(* IEC 61131-3 sources: IRIS-Project/LASAL CONTROL SOFTWARE/LasalProject_2025_09_25/Runtime/%LASALAPPDATA%/Runtime/Library/Loader/Source/code (part 3) *)

  IF SramdiskNotWrittenAtPowerDown() THEN
		DEBUGLOG0("%010d error: sramdisk was not written at power-down");
    _s_ram_hptr^.DataValid$UINT := 0;
    sramErrorCode := EC_SRAMDISK_NOT_WRITTEN_AT_POWER_DOWN;
    LogSramError();
  END_IF;

	IF isRamfileDatUsed THEN
		// Das RAMFILE.DAT auf pRamFile einlesen
		IF SramLoadFile() <> 0 THEN
			_s_ram_hptr^.DataValid$UINT := 0;
			sramErrorCode := EC_LOADFILE_ERR;
			LogSramError();
		ELSIF IsVortex() = FALSE & WasRemoveableMediaChanged() THEN
			DEBUGLOG0("%010d error: detected media change, ramfile.dat not usable, marking sram as invalid");
			_s_ram_hptr^.DataValid$UINT := 0;
		END_IF;
	END_IF;

  fDoNotReportErrors := 0;
  IF GetSramReorgFlag() & ((_s_ram_hptr^.DataValid AND 16#FF000000) = 16#80000000) THEN
    // Wenn das Reorg-Flag im DataValid Feld gesetzt ist, dann heißt das, daß
    // ein Reorg Vorgang unterbrochen wurde, nachdem eine File Kopie angelegt
    // wurde. In so einem Fall wird keine Fehlermeldung generiert.
    fDoNotReportErrors := 1;
  END_IF;

	IF GetSramReorgFlag() THEN
		fReorgSram := 1;
	END_IF;
	wasValid := CHK_S_RAM(fDoNotReportErrors);
	IF GetSramReorgFlag() THEN
		IF wasValid THEN

			// gültigen SRAM Inhalt auf Files kopieren
			rc := MakeSramKopie(#errCode);
			IF rc = 0 THEN

				// Der SRAM Inhalt befindet jetzt als Kopie in den Files.
				// Es wird jetzt als ungültig gekennzeichnet und durch den Aufruf von CHK_S_RAM
				// wird das SRAM noch einmal mit 0 initialisiert.
				DEBUGLOG0("%010d MakeSramKopie succeeded, marking sram as invalid");

				_s_ram_hptr^.DataValid$UINT := 0;
        // Das Reorg-Flag setzen. Wenn dieses Flag gesetz ist, dann heisst das, daß
        // das SRAM zwar ungültig ist, aber eine gültige Kopie im File existiert.
        // In diesem Fall (ungültige SRAM, gültige Kopie im File) wird kein SRAM
        // Fehler gemeldet.
        _s_ram_hptr^.DataValid := (_s_ram_hptr^.DataValid AND 16#00FFFFFF) OR 16#80000000;

        // Der folgende Aufruf von CHK_S_RAM bewirkt, daß das SRAM neu initilisiert
        // wird (weil DataValud 0 ist).
				fReorgSram := 1;
				CHK_S_RAM(fDoNotReportErrors := 1);
        // Reorg-Flag muss hier noch einmal gesetzt werden, da CHK_S_RAM den
        // ganzen Header auf 0 setzt.
        _s_ram_hptr^.DataValid := (_s_ram_hptr^.DataValid AND 16#00FFFFFF) OR 16#80000000;

			ELSE
				DEBUGLOG2("%010d MakeSramKopie failed, rc=%d, errCode = 0x%X" , rc$UDINT, errCode$UDINT);
			END_IF;

		//ELSIF !!WasRemoveableMediaChanged() THEN
    ELSE
			_s_ram_hptr^.DataValid$UINT := 0;
            // Der folgende Aufruf von CHK_S_RAM bewirkt, daß das SRAM neu initilisiert
            // wird (weil DataValid 0 ist). Das ist notwendig, damit in der MAT die
			// durch SRAM_MARKMemory belegten Bereiche wieder freigegeben werden.
			// (SRAM_MARKMemory wurde in CHK_S_RAM aufgerufen, um die vorhandenen
			// SRAM Einträge als belegt zu markieren).
			fReorgSram := 1;
			CHK_S_RAM(fDoNotReportErrors := 1);

			// Das SRAM war ungültig, durch das Setzen des Flags fReorgSram wird
			// versucht, auf Daten von einer früheren Kopie zurückzugreifen.
			fReorgSram := 1;
			DEBUGLOG0("%010d MakeSramKopie: no copy created, because sram is not valid");
		END_IF;
	END_IF;

	CLEAR_LASTENTRY();

END_FUNCTION

//------------------------------------------------------------------------
// S-Ram Initialisieren und ggf alte formate konvertieren (aus active.dat)
//-------------------------------------------------------------------------
// Bei aufruf hat das BS schon in  "_S_RAM_Hptr"  einen pointer auf den S-Ram-Descriptor
// Descriptor eingetragen (oder auch nicht. ein altes system hat dort 0 stehen
//
// Logik : a) _S_RAM_Hptr hat einen gültigen pointer.
//				Wenn der eintrag genutzte länge > 0 ist gelten diese daten
//				Wenn der eintrag genutzte länge = 0 ist, suchen wir eine Active.dat
//
// 06.03.04
// wenn C-IPC konvertieren auf neues format
// es stehen nur noch die Daten im Ram der Rest ist in einem File
// so sparen wir pro eintrag 12 Byte !!!
//
//

FUNCTION S_RAM_INIT

VAR_OUTPUT
	ret_code 		: CONFSTATES;
END_VAR

VAR
	ActiveDatHandle  :DINT;
	DateiKopf     : DatKopf;
	OneRecord     : Eintrag;
	RecNr		  : UDINT;
	I			  : DINT;
	PtChar		  : ^CHAR;
	PtxNextRAM	  : ^XRamCell;
	ptxRamHead	  : ^XRAMHDR;
	RelAdress	  :  UDINT;
  formatChanged : BOOL;
  initCnt : UDINT;
	gotMemory : BOOL;
END_VAR

  if !!hasSram then
    ret_code:=C_OK;
    return;
  end_if;

  CONVERT_SRAM();

	// das erstellen wir automatisch
  if _rtosversion > 16#537 then
    if LSLFILE_IsInstalled then
      // Das Direktory für die File Daten erstellen
      OS_FILE_CREATEDIR("C:\FData");
    end_if;
  end_if;

  ret_code:=C_OK;
  initCnt := 0;
Brutal_start:
  initCnt += 1;

//---------------------------------------
// Wenn Neues BS ist der Ptr ungleich 0
//---------------------------------------

  IF _S_RAM_Hptr <> 0 then      // Diesen Pointer gibt es seit a.m mit pranz und gradl am 2.2.2002 vergangenheitsbewältigung gemacht hat

    if (_S_RAM_Hptr^.DataLength <= maxSramSize) then
      SRAM_STARTUP(_S_RAM_Hptr^.DataLength , 1);
    else
      SRAM_STARTUP(maxSramSize, 1);  // SRAM begrenzen
    end_if;

    //------------------------------------------------------
    // wenn jungfräulich, test ob alte active.dat vorhanden
    //------------------------------------------------------
    IF _S_RAM_Hptr^.UsedData = 0 then

      //-- Neues _SRAM Löschen ---

      // Der Aufruf dieser Funktion bewirkt, dass auch bei gelöschtem Sram
      // das File sernum.dat, wo die Seriennummer gespeichert ist, erstellt wird.
      WasRemoveableMediaChanged();

      RelAdress:=InitXramBlockEx(#gotMemory);
      IF gotMemory THEN
        ptxRamHead:= _S_RAM_Hptr^.DataStart+RelAdress;
        PtxNextRam:=#ptxRamHead^.aData[0];

        // active.dat nur möglich wenn filesystem vorhanden

        IF (LSLFILE_IsInstalled) THEN

          ActiveDatHandle:=OS_FILE_OPEN("c:\active.dat",0,16#000);

          // das file ist gefunden -> konvertieren
          IF ActiveDatHandle > 0 THEN
            OS_FILE_READ(ActiveDatHandle, #DateiKopf.signi[0], sizeof(DateiKopf));
            IF DateiKopf.NrRec <> 0 then  // #FA wenn keine eintraege ende  (gibt es auch)
              FOR RecNr:= 0 to DateiKopf.NrRec -1 do
                // -- GUID LESEN
                OS_FILE_READ(ActiveDatHandle,#OneRecord.myguid[0],sizeof(Eintrag.myguid));
                // -- NAMEN LESEN

                PtCHar:=#OneRecord.Name[0];
                FOR I:= 0 to SIZEOF(Eintrag.Name) -1 do
                  OS_FILE_READ(ActiveDatHandle,PtCHar,1);
                  if PtChar^ =0 then
                    GOTO GOTNAME;
                  elsif PtChar^ = '.' then
                    PtChar^:=0;
                  end_if;
                  PtCHar+=1;
                END_FOR;

                // ERROR NAME TO LONG !!!!

                ret_code:=C_OUTOF_NEAR;
                OS_FILE_CLOSE(ActiveDatHandle);
                GOTO	Brutal_ende;

              //...........................
              // Der Name ist eingelesen !
              //...........................

              GOTNAME:

                // wenn block voll, neuen block erzeugen & Verkettung herstellen

                if ptxRamHead^.udEntries = X_RAM_CELLS	then
                  RelAdress:=IniNewRamBlock(PtxNextRam);
                  If Reladress <> 0 then
                    ptxRamHead:= _S_RAM_Hptr^.DataStart+RelAdress;
                    PtxNextRam:=#ptxRamHead^.aData[0];
                    // Kein platz mehr im RAM !!!
                  else
                    ret_code:=C_OUTOF_NEAR;
                    OS_FILE_CLOSE(ActiveDatHandle);
                    GOTO	Brutal_ende;
                  end_if;
                end_if;

                // Daten und Sizeof daten lesen

                OneRecord.CRC:=CRC32(#OneRecord.Name[0]);

                OS_FILE_READ(ActiveDatHandle,#OneRecord.Data,2*4);

                // Wenn Len > 0 dann ist es eine RAMEX falls es eine RAMEX mit 0 ist
                // kommt das später beim Instanzieren dran

                IF OneRecord.Len <> 0 then
                  RelAdress$UDINT:= (SRAM_GetMemory(OneRecord.Len$UDINT))$UDINT;
                  If Reladress <> 0 then

                    PtxNextRam^.udType:=IsXram$UDINT+RelAdress$UDINT;
                    OS_FILE_READ(ActiveDatHandle,_S_RAM_Hptr^.DataStart+RelAdress,OneRecord.Len$UDINT);
                    // in the data HIGH Part is the real length
                    // in the lo part the allocated length
                    OneRecord.Data$UDINT := OneRecord.Len$UDINT SHL 16;
                    OneRecord.Data$UDINT := OneRecord.Data$UDINT OR  SRAM_GET_ALLOCATED(OneRecord.Len$UDINT);
                  end_if;

                ELSE
                  PtxNextRam^.udType:= 0;
                END_IF;

                PtxNextRam^.udCRC32:=OneRecord.CRC;
                PtxNextRam^.udData$UDINT:=OneRecord.Data$UDINT;
                PtxNextRam^.udChk$UDINT:=OneRecord.Data$UDINT+OneRecord.CRC+(PtxNextRam^.udType$UDINT AND 16#00ffFFFF);
                PtxNextRam^.udType:=PtxNextRam^.udType or RamValid;  // VALID RAM LOCATION

                ptxNextRam+=SIZEOF(xRamCell);
                ptxRamHead^.udEntries+=1;
                ptxRamHead^.udChk:=NOT ptxRamHead^.udEntries;

              END_FOR;
            END_IF;
            OS_FILE_CLOSE(ActiveDatHandle);
            S_RAM_INIT_I();

          // keine active.dat vorhanden  und neues system und dateisystemvorhanden .
          //--> Speicher Initialisieren
          ELSE
            S_RAM_INIT_I();
          END_IF;

        // Kein filesystem vorhanden & keine daten: jungfräulich, initialisieren
        // oder das alte Format konvertieren !
        // muss eigentlich Eine 386 sein ??

        ELSE
          // #FA
          // wir versuchen die alten daten auch zu konvertieren aber nur einmal
          if aRamHdr.udEntries <> 0 then
            if aRamHdr.udEntries = NOT aRamHdr.udChk then
              if aRamHdr.udEntries < 1000 then // sicherheit
                // schleife für die konvertierung bilden !!!
                for RecNr:=0 to (aRamHdr.udEntries-1) do

                  // wenn block voll, neuen block erzeugen & Verkettung herstellen
                  if ptxRamHead^.udEntries = X_RAM_CELLS	then
                    RelAdress:=IniNewRamBlock(PtxNextRam);
                    If Reladress <> 0 then
                      ptxRamHead:= _S_RAM_Hptr^.DataStart+RelAdress;
                      PtxNextRam:=#ptxRamHead^.aData[0];
                    // Kein platz mehr im RAM !!!
                    else
                      ret_code:=C_OUTOF_NEAR;
                      GOTO	Brutal_ende;
                    end_if;
                  end_if;

                  // check if chk is o.k.
                  if aRamHdr.aData[RecNr].udChk = aRamHdr.aData[RecNr].udCRC32 + aRamHdr.aData[RecNr].udData then
                    PtxNextRam^.udCRC32:=aRamHdr.aData[RecNr].udCRC32;
                    PtxNextRam^.udData$UDINT:=aRamHdr.aData[RecNr].udData;
                    PtxNextRam^.udChk$UDINT:=aRamHdr.aData[RecNr].udChk;

                    PtxNextRam^.udType:=PtxNextRam^.udType or RamValid;  // VALID RAM LOCATION

                    ptxNextRam+=SIZEOF(xRamCell);
                    ptxRamHead^.udEntries+=1;
                    ptxRamHead^.udChk:=NOT ptxRamHead^.udEntries;
                  end_if;

                end_for;
              end_if;
            end_if;
            aRamHdr.udEntries :=0;
            aRamHdr.udChk :=0;
          end_if;

          S_RAM_INIT_I();
        END_IF;
      ELSE // gotMemory
        IF !!isRamfileDatUsed THEN
          // Bei SRAM Format 1 muss auf jeden Fall der xRamHdr Platz haben
          LDR_outOfSramMem := TRUE;
        END_IF;

        S_RAM_INIT_I();
      END_IF;

    //--- ES SIND DATEN VORHANDEN, TESTEN !!! ---

    ELSE
      S_RAM_INIT_I();
    END_IF;

  //------------------------------------
  // ALTES FORMAT (kein Ptr auf ram vorhanden)
  //------------------------------------
  else
    ret_code:=C_OUTOF_NEAR;
  END_IF;
Brutal_ende:

  IF loaderRamexError THEN
    IF isSramNewOrCleared THEN
      DEBUGLOG0("%010d-resetting sram content due to a detected new or cleared sram");
    ELSE
      DEBUGLOG0("%010d-resetting sram content due to a detected error");
    END_IF;
    LDR_outOfSramMem := FALSE;
    _s_ram_hptr^.UsedData := 0;
    _s_ram_hptr^.DataStart^.udEntries := 0;
    _s_ram_hptr^.DataStart^.udChk:=NOT _s_ram_hptr^.DataStart^.udEntries;
    IF GetRamfileDatUsedFlag(#formatChanged) THEN
      _s_ram_hptr^.DataValid := 0x20001;
    ELSE
      _s_ram_hptr^.DataValid := 0x00001;
    END_IF;
    IF pRamFile THEN
      pRamFile^.udEntries :=  0;
      pRamFile^.uiChange  :=  16#1234;	// änderung eintragen wir speicher hier gleich
    END_IF;
    SramSaveFile();

    // DS2589, 02.02.182, 9.5.2016:
    // Eine möglicherweise von früher noch vorhandene Sram-Kopie (vom Reorganisieren)
    // wird gelöscht, damit im Fall einer gesetzten SRAM_CONTINUE_ON_ERROR Umgebungsvariable
    // das Sram mit den Init-Werten und nicht mit den Werten aus der Kopie initialisiert wird.
    DeleteSramKopie();

    IF (!!bSramContinueOnError & !!isSramNewOrCleared) | (initCnt > 1) THEN
      ret_code:=C_OUTOF_NEAR;
    ELSIF formatChanged THEN
      // Wenn das Format geändert wurde, dann muss noch einmal initialisiert
      // werden (es ist z.B. die Größe der MAT vom Format abhängig).
      loaderRamexError := 0;
      GOTO Brutal_start;
    END_IF;
  END_IF;

END_FUNCTION

// Löscht im alten Format in der letzten Zelle des ersten Blocks den im Element
// udType (in den untersten 20 Bits) gespeicherten Merker für die letzte gefundene
// Ramzelle. Dieser Merker wird von der Funktion Find_sRam_I zum Zwischenspeichern
// des Block-Index und Zell-Offsets der zuletzt gefundenen Zelle verwendet.
// Damit wird die Suche schneller, wenn Find_sRam_I nicht jedesmal von vorne
// zu suchen beginnt, sondern dort wo sie den letzten Eintrag gefunden hat.
//
// Im neuen Format (mit ramfile.dat) wird dieser Merker nicht verwendet.
FUNCTION CLEAR_LASTENTRY
VAR
  pRamCell : ^XRamCell;
END_VAR;

  IF (_S_RAM_Hptr^.DataValid SHR 16) < 2 &  _s_ram_hptr^.DataLength >= SIZEOF(XRAMHDR) THEN
    // altes Format
    pRamCell := #_S_RAM_Hptr^.DataStart^.aData[X_RAM_CELLS];
    pRamCell^.udType := pRamCell^.udType AND 16#FFF0_0000;
  END_IF;

END_FUNCTION

// loescht alle Einträge
FUNCTION ClearEntrys

	pRamFile^.udEntries   := 0;
	pRamFile^.CRC32       := 0;
	pRamFile^.pLastEntry  := 0;

END_FUNCTION

#define READ_COMPLETE_RAMFILEDAT

// Wenn das Sram im RAM liegt mit einem Backup auf SD Karte (Edge-CPUs),
// dann wird in dieser Funktion der Sram-Inhalt auf die SD Karte gesichert.
FUNCTION FlushSramToDisk
VAR
  pSrd : ^OS_SRAMDISK;
END_VAR

  OS_CILGet("SRAMDISK", #pSrd$void);
  IF (pSrd <> NIL) & (pSrd^.udVersion >= 2) THEN
    SRAMDISK_COMMIT(pSrd);
#ifdef _LSL_TARGETARCH_X86
    // SA26191,DS2087: Workaround für einen OS-Fehler bei ETVEdge Plattformen:
    // Interrupts sind nach Aufruf von SRAMDISK_COMMIT gesperrt, wenn fullCopyAtPowerdown gesetzt ist.
    // Die Interrupts werden hier wieder freigegeben.
    IF _RtOSVersion < 16#9000 THEN
      STI();
    END_IF;
#endif
  END_IF;

END_FUNCTION

// funktion schreibt daten auf Flash falls verson C-IPC +
// die Version > 2 ist und sich auch was geändert hat !! in diesem File
FUNCTION GLOBAL SramSaveFile
VAR
	Handle : DINT;
	CRC32  : UDINT;
	aXFileHdr_Hdr : XFILEHDR_HDR;
	pCopy  : ^XFILEHDR;
	rc     : UDINT;
	bytes2Write	 : UDINT;
	bytes2Read   : UDINT;
  allocSize : UDINT;
  att : UDINT;
END_VAR

  if !!hasSram then
    return;
  end_if;

	// test auf C-IPC
	if isRamfileDatUsed then
 	  // test auf pointer vorhanden und version groesser 1
	  if (_S_RAM_Hptr <> NIL) & ((_S_RAM_Hptr^.DataValid shr 16) > 1) then

      if pRamFile^.uichange <> 16#1234 then
        // Wenn keine Änderung war und noch kein RamFile.dat existiert (neuer CIPC),
        // dann wird pRamFile^.uichange auf 16#1234 gesetzt. Dadurch wird das Anlegen
        // eines (leeren) RamFile.dat erzwungen.
        Handle:=OS_FILE_OPEN("c:\RamFile.dat",0,16#000);	// read-only
        if handle >= 0 then
          OS_FILE_CLOSE(handle);
        else
          pRamFile^.uichange := 16#1234;
        end_if;
      end_if;

      // test ob auch sich was geändert hat
      if pRamFile^.uichange = 16#1234 then
        // Ab 1.1.27 wird das SRAM bei jedem Start reorganisiert.
        // Die pRamFile Struktur wird immer neu aufgebaut, d.h. uichange hat
        // dann immer den Wert 16#1234 weil immer Änderungen gemacht werden.
        // Jetzt kann es aber sein, daß die Struktur gleich geblieben ist (wenn sich
        // die Checksumme und udEntries nicht geändert hat). Wenn das der Fall ist, dann
        // wird uichange auf 0 gesetzt, damit das RAMFILE.DAT nicht unnötigerweise
        // neu erstellt wird.

        // Checksumme rechnen
  #ifdef READ_COMPLETE_RAMFILEDAT
        CRC32 := CALC_RAMFILE_DAT_CRC(pRamFile);
  #else
        CRC32:=CRC32_Buffer(#pRamFile^.aData,pRamFile^.udEntries * SIZEOF(XFileCell));
  #endif
        // Checksumme aus dem File einlesen und vergleichen
        handle := OS_FILE_OPEN("c:\RamFile.dat", 0, 0);		// 0 = read only
        IF handle > 0 THEN
          rc := OS_FILE_READ(handle, #aXFileHdr_Hdr, SIZEOF(aXFileHdr_Hdr));
          IF rc = SIZEOF(XFileHdr_Hdr) THEN
            IF (aXFileHdr_Hdr.CRC32 = CRC32) & (aXFileHdr_Hdr.udEntries = pRamFile^.udEntries) THEN
              pRamFile^.uichange := 0;
              DEBUGLOG2("%010d-SramSaveFile: no need to write to ramfile.dat (crc32=0x%08X and udEntries=%d are still the same)", CRC32, pRamFile^.udEntries);
            END_IF;
          END_IF;
          OS_FILE_CLOSE(handle);
        END_IF;
      end_if;

      if pRamFile^.uichange = 16#1234 then

        pRamFile^.CRC32 := CRC32;

				// RAMFILE.DAT auf RAMFILE.BAK kopieren
        Handle:=OS_FILE_OPEN("c:\RamFile.dat",0,16#000);
	      if handle >= 0 then
          allocSize := XFILEHDR.adata + X_FILE_CELLS_2 * SIZEOF(XFileCell);
     			pCopy := (_alloc_resize_LDR(allocSize))$^XFILEHDR;
		      if pCopy <> NIL then
						bytes2Read := allocSize;
	     			rc := OS_FILE_READ(Handle, pCopy, bytes2Read);
		        OS_FILE_CLOSE(handle);
						if rc < 0 then
							DEBUGLOG2("%010d-SramSaveFile: error reading ramfile.dat, bytes2read=%d, rc=%d", bytes2read, rc);
						else
		          handle:=OS_FILE_OPEN("c:\RamFile.bak",2,ATT_CREATE);
							if handle >= 0 then
								bytes2Write := rc;
			 					rc := FileWrite(handle, pCopy, bytes2Write)$UDINT;
								if rc <> bytes2Write then
									DEBUGLOG2("%010d-SramSaveFile: error writing ramfile.bak, bytes2write=%d, rc=%d", bytes2Write, rc);
								else
									DEBUGLOG1("%010d-SramSaveFile: ramfile.dat copied into ramfile.bak (%d bytes)", rc);
								end_if;
				 				OS_FILE_CLOSE(handle);
							else
								DEBUGLOG1("%010d-SramSaveFile: could not open ramfile.bak, rc=%d", handle$UDINT);
							end_if;
	          end_if;
	     		  _free(pCopy);
					else
					  DEBUGLOG1("%010d-SramSaveFile: could not allocate enough memory (%d)", allocSize$UDINT);
		        OS_FILE_CLOSE(handle);
	        end_if;
	   		end_if;

        // den Inhalt von pRamFile ins File RAMFILE.DAT schreiben
        if pRamFile^.udEntries > X_FILE_CELLS then
          bytes2Write := XFILEHDR.adata + X_FILE_CELLS_2 * SIZEOF(XFileCell);
        else
          bytes2Write := XFILEHDR.adata + X_FILE_CELLS * SIZEOF(XFileCell);
        end_if;
        if bytes2Write <> LDR_allocated_XFileSize then
          att := ATT_CREATE_ALWAYS;
        else
          att := ATT_CREATE;
        end_if;

        handle:=OS_FILE_OPEN("c:\RamFile.dat", 2, att);
        if Handle >= 0 then
          rc := FileWrite(handle, pRamFile, bytes2Write)$UDINT;
          if rc <> bytes2Write then
            DEBUGLOG2("%010d-SramSaveFile: error writing ramfile.dat, bytes2write=%d, rc=%d", bytes2Write, rc);
            SramError();
          else
            DEBUGLOG3("%010d-SramSaveFile: data written to ramfile.dat (%d bytes, crc32=0x%X), udEntries=%d", rc, pRamFile^.CRC32, pRamFile^.udEntries);
            // Wenn das Sram im RAM liegt mit einem Backup auf SD Karte (Edge-CPUs),
            // dann wird nach dem Ändern der ramfile.dat der Sram-Inhalt auf die SD Karte
            // geschrieben. Damit ist ramfile.dat und Sram konsistent, auch für den Fall dass
            // beim Abschalten das Sram nicht mehr auf die SD Karte geschriben wird.
            FlushSramToDisk();
            pRamFile^.uichange := 0;
          end_if;
          OS_FILE_CLOSE(handle);
        else
          DEBUGLOG1("%010d-SramSaveFile: could not open ramfile.dat, rc=%d", handle$UDINT);
          Trace_ERR("SAVE OF RamFile not possible (Disk full??)");
          LSLCLI_LoaderTracePrint("SAVE OF RamFile not possible (Disk full??)", 12);
          SramError();
        end_if;

        // ramfile.bak ungültig machen, nachdem ramfile.dat erstellt worden ist
        InvalidateRamfileBak();

      end_if;
    end_if;
	end_if;
END_FUNCTION

// ------------------------------------------
//   laden des File von C-IPC in Speicher
// ------------------------------------------
// das file ist 192k /4 Byte (je Eintrag im S-RAM) * 12 byte (je Eintrag im File)
// groß = 576 k Byte
// die RamEx bleibt so wie alt
// udCRC32    (4 Byte)
// udType     (4 Byte)
// udpRelSram (4 Byte)

FUNCTION SramLoadFile
VAR_OUTPUT
	result : UDINT;
END_VAR
VAR
	Handle : DINT;
	CRC32  : UDINT;
	rc     : UDINT;
	bytes2Read   : UDINT;
	fileSize   : UDINT;
  udEntries_file  : UDINT;
  nCellsAlloc : UDINT;
  allocSize : UDINT;
END_VAR
  result := 16#FFFFFFFF;

  // Die Anzahl der benötigten Zellen ist erst nach dem Lesen des Ramfile.dat
  // bekannt, da aber nachfolgender Code davon ausgeht, dass pRamfile <> NIL ist, wird
  // hier einmal mit X_FILE_CELLS allokiert. Ggf. wird das dann noch vergrößert.
  nCellsAlloc := X_FILE_CELLS;
  allocSize := XFILEHDR.adata + nCellsAlloc * SIZEOF(XFileCell);
	pRamFile := _alloc_resize_LDR(allocSize)$^XFILEHDR;
  if pRamFile <> NIL then
    LDR_allocated_XFileCells := nCellsAlloc;
    LDR_allocated_XFileSize := allocSize;
    ClearEntrys();
  end_if;

  Handle := OS_FILE_OPEN("c:\RamFile.dat",0,0);
  if Handle < 0 then
    DEBUGLOG1("%010d-SramLoadFile: could not open ramfile.dat, rc=%d", handle$UDINT);
    SramError();
    return;
  end_if;
  rc := OS_FILE_READ(Handle, #udEntries_file, SIZEOF(udEntries_file));
  if rc <> SIZEOF(udEntries_file) then
    DEBUGLOG1("%010d-SramLoadFile: could not read udEntries_file from ramfile.dat, rc=%d", rc);
    SramError();
    return;
  end_if;
  OS_FILE_CLOSE(handle);

  if udEntries_file > X_FILE_CELLS & pRamFile <> NIL then
    nCellsAlloc := X_FILE_CELLS_2;
    allocSize := XFILEHDR.adata + nCellsAlloc * SIZEOF(XFileCell);
   	pRamFile := _realloc_LDR(pRamFile, allocSize)$^XFILEHDR;
  end_if;

  if pRamFile <> NIL then
    LDR_allocated_XFileCells := nCellsAlloc;
    LDR_allocated_XFileSize := allocSize;

    ClearEntrys();

    // try to open file
    Handle:=OS_FILE_OPEN("c:\RamFile.dat",0,0);
	  if Handle > 0 then
	 // file ist da laden
#ifdef READ_COMPLETE_RAMFILEDAT
			bytes2Read := allocSize;
			rc := OS_FILE_READ(Handle, pRamFile, bytes2Read);
#else
			rc := OS_FILE_READ(Handle, pRamFile, SIZEOF(XFILEHDR.udEntries));
      if rc = SIZEOF(XFILEHDR.udEntries) then
			  bytes2Read := XFILEHDR.adata + pRamFile^.udEntries * SIZEOF(XFileCell) - SIZEOF(XFILEHDR.udEntries);
			  rc := OS_FILE_READ(Handle, pRamFile + SIZEOF(XFILEHDR.udEntries), bytes2Read);
      end_if;
#endif
	    OS_FILE_CLOSE(handle);
      fileSize := XFILEHDR.adata + pRamFile^.udEntries * SIZEOF(XFileCell);
			if rc < 0 then
				DEBUGLOG1("%010d-SramLoadFile: error reading ramfile.dat, no header information, rc=%d", rc);
				SramError();
			elsif rc <> bytes2Read then
				DEBUGLOG3("%010d-SramLoadFile: error reading ramfile.dat, fileSize=%d, bytes2Read=%d, rc=%d", fileSize, bytes2Read, rc);
				SramError();
			else
	      // file im Speicher CRC rechnen
	      pRamFile^.uiChange :=0;				// keine Änderung
	      pRamFile^.pLastEntry :=0;				// und von anfang an
#ifdef READ_COMPLETE_RAMFILEDAT
	      CRC32 := CALC_RAMFILE_DAT_CRC(pRamFile);
#else
	      CRC32:=CRC32_Buffer(#pRamFile^.aData,pRamFile^.udEntries * SIZEOF(XFileCell));
#endif

	      if CRC32 = pRamFile^.CRC32 then
	        // file im speicher CRC = o.k. wir belegen den Speicher
	        if ((pRamFile^.udEntries <> 0) & (pRamFile^.udEntries <= X_FILE_CELLS_2)) then
						DEBUGLOG2("%010d-SramLoadFile: data read from ramfile.dat (%d bytes), udEntries=%d", rc, pRamFile^.udEntries);
	          result:=0;
	        else
						if pRamFile^.udEntries > X_FILE_CELLS_2 then
					  	DEBUGLOG1("%010d-SramLoadFile: invalid udEntries (%08X)", pRamFile^.udEntries);
						  SramError();
						else
							result := 0;
						end_if;
						ClearEntrys(); // 0 oder zu viele einträge
  	      end_if;
	      else
					DEBUGLOG2("%010d-SramLoadFile: invalid crc32 (calc:0x%08X, file:0x%08X)", CRC32, pRamFile^.CRC32);
					// die CRC ist falsch

					Handle := OS_FILE_OPEN("c:\RamFile.er1",2,ATT_CREATE);
					FileWrite(handle,pRamFile, allocSize);
					OS_FILE_CLOSE(handle);

          // wir nehmen das BAK falls vorhanden
          Handle:=OS_FILE_OPEN("c:\RamFile.bak",2,ATT_READ_WRITE);
          if Handle > 0 then
            OS_FILE_CLOSE(handle);
            OS_FILE_DELETE("c:\RamFile.dat");
            OS_FILE_RENAME("c:\RamFile.bak", "c:\RamFile.dat");
            _free(pRamFile);			// wird nochmal gemacht !!
            result:=SramLoadFile();	// rekursion !!
          end_if;
	      end_if;
	    end_if;
	  else
			DEBUGLOG1("%010d-SramLoadFile: could not open ramfile.dat, rc=%d", handle$UDINT);
			SramError();
	  end_if;
  end_if;

	IF result <> 0 THEN
   		DEBUGLOG1("%010d-SramLoadFile failed, rc=%d", result);
	END_IF;

END_FUNCTION

//------------------------------------------------------------------------------
// AlarmSramError
//------------------------------------------------------------------------------
FUNCTION AlarmSramError
VAR_INPUT
  param : DINT;
END_VAR
	IF (pSramAlarmSvrCh = NIL) & ( (OPS.SysState = C_RUNRAM) | (OPS.SysState = C_RUNROM) ) THEN
		_LookUpEmbed_C(SRAMALARM_SVR_NAME, #pSramAlarmSvrCh, NIL);
	END_IF;
	IF pSramAlarmSvrCh <> NIL THEN
		ESI := pSramAlarmSvrCh;
		pSramAlarmSvrCh^.pMeth^.pWr$M_WR_DIRECT(param);
	END_IF;
END_FUNCTION
//------------------------------------------------------------------------------
// SramError
//------------------------------------------------------------------------------
FUNCTION SramError
	IF loaderRamexError = 0 THEN
    IF isSramNewOrCleared THEN
		  TRACE("New or cleared SRAM detected, see c:\sysmsg\event19.log. Resetted SRAM.");
      LSLCLI_LoaderTracePrint("New or cleared SRAM detected, see c:\sysmsg\event19.log. Resetted SRAM.", 12);
    ELSIF bSramContinueOnError THEN
		  TRACE_WARN("Error in SRAM, see c:\sysmsg\event19.log. Resetted SRAM.");
      LSLCLI_LoaderTracePrint("Error in SRAM, see c:\sysmsg\event19.log. Resetted SRAM.", 12);
    ELSE
		  TRACE_WARN("Error in SRAM, see c:\sysmsg\event19.log. Resetted SRAM, project must be restarted");
      LSLCLI_LoaderTracePrint("Error in SRAM, see c:\sysmsg\event19.log. Resetted SRAM, project must be restarted", 12);
    END_IF;
	END_IF;
	loaderRamexError := 1;
END_FUNCTION
//------------------------------------------------------------------------------
// LogSramError
//------------------------------------------------------------------------------
FUNCTION LogSramError
	IF sramErrorCode = 4 THEN
		// Der Fehlercode 4 kommt zustande, wenn ein RAMFILE.DAT mit udEntries = 0
		// vorgefunden wird.
		// pr:
		//	Meiner Meinung nach ist das kein Fehler, daher wird hier keine Meldung
		//  ausgegeben.
		//  Es wird aber trotzdem der Code für die Fehlerbehandlung durchlaufen, weil
		//  ich nicht weiss wie der ganze Assemblercode auf udEntries = 0 reagieren würde.
		RETURN;
	END_IF;
	DEBUGLOG1("%010d-SramError, errorCode=%08X", sramErrorCode);
	IF _S_RAM_Hptr THEN
		DEBUGLOG1("%010d             Version    = %08X" , _S_RAM_Hptr^.Version);
		DEBUGLOG1("%010d             DataStart  = %08X" , _S_RAM_Hptr^.DataStart$UDINT);
		DEBUGLOG1("%010d             DataLength = %08X" , _S_RAM_Hptr^.DataLength);
		DEBUGLOG1("%010d             UsedData   = %08X" , _S_RAM_Hptr^.UsedData);
		DEBUGLOG1("%010d             DataValid  = %08X" , _S_RAM_Hptr^.DataValid);
		IF _S_RAM_Hptr^.DataStart THEN
			DEBUGLOG1("%010d             udEntries  = %08X" , _S_RAM_Hptr^.DataStart^.udEntries);
			DEBUGLOG1("%010d             udChk      = %08X" , _S_RAM_Hptr^.DataStart^.udChk);
		END_IF;
	END_IF;
	SramError();
END_FUNCTION
//------------------------------------------------------------------------------
// LogSramRamexError
//------------------------------------------------------------------------------
FUNCTION __CDECL LogSramRamexError
VAR_INPUT
	pXramCell : ^XRamCell;
END_VAR
	DEBUGLOG1("%010d-RamexError, cellAddr = %08X" , pXramCell$UDINT);
	DEBUGLOG1("%010d             udChk    = %08X" , pXramCell^.udChk);
	DEBUGLOG1("%010d             udCRC32  = %08X" , pXramCell^.udCRC32);
	DEBUGLOG1("%010d             udData   = %08X" , pXramCell^.udData);
	DEBUGLOG1("%010d             udType   = %08X" , pXramCell^.udType);
	SramError();
END_FUNCTION
//------------------------------------------------------------------------------
// LogSramChk
//------------------------------------------------------------------------------
FUNCTION LogSramChk
	DEBUGLOG0("%010d-checking Sram");
END_FUNCTION
//------------------------------------------------------------------------------
// SramCheckerInit
//------------------------------------------------------------------------------
FUNCTION SramCheckerInit
	fileCellChkIdx := 0;
END_FUNCTION

#ifdef CYCLIC_SRAM_CHECK
#define CELLMASK_VALID      0x80000000
#define CELLMASK_USED       0x40000000
#define CELLMASK_CELLTYPE   0x3C000000
#define CELLMASK_RAMEXADR   0x00FFFFFF

#define CELLTYPE_RAM        0x00000000
#define CELLTYPE_RAMEX      0x30000000

FUNCTION SramCheckV1
VAR
  pHdr : ^XRAMHDR;
  sramStart : pVoid;
  sramEnd : pVoid;
  pCellEnd : ^XRamCell;
  pCell : ^XRamCell;
  cellChksum : UDINT;
END_VAR

  sramStart := _S_RAM_Hptr^.dataStart;
  sramEnd := sramStart + _S_RAM_Hptr^.dataLength;
  pHdr := _S_RAM_Hptr^.dataStart;

  WHILE ((pHdr >= sramStart) & (pHdr < sramEnd)) DO

    IF pHdr^.udEntries > X_RAM_CELLS + 1 THEN
  		sramErrorCode := EC_INV_BLK_ENTRIES;
      SramError();
      AlarmSramError(pHdr$DINT);
    END_IF;
    IF (pHdr^.udEntries XOR pHdr^.udChk) <> 16#FFFFffff THEN
  		sramErrorCode := EC_INV_BLK_CHKSUM;
      SramError();
      AlarmSramError(pHdr$DINT);
    END_IF;

    pCell := #pHdr^.aData[0];
    pCellEnd := #pHdr^.aData[pHdr^.udEntries];
    WHILE pCell < pCellEnd DO

      IF pCell^.udType AND CELLMASK_VALID THEN
        IF pCell^.udType AND CELLMASK_CELLTYPE AND CELLTYPE_RAMEX THEN
          cellChksum := pCell^.udData + pCell^.udCRC32 + (pCell^.udType AND CELLMASK_RAMEXADR);
        ELSE
          cellChksum := pCell^.udData + pCell^.udCRC32;
        END_IF;
        IF cellChksum <> pCell^.udChk THEN
      		sramErrorCode := EC_INV_CELL_CHKSUM;
          SramError();
          AlarmSramError(pCell$DINT);
        END_IF;
      END_IF;

      pCell += sizeof(XRamCell);
    END_WHILE;

    IF pCell = #pHdr^.aData[X_RAM_CELLS] THEN
      // Block war zur Gänze gefüllt
      // prüfen, ob die 501. Zelle auf einen weiteren Block zeigt
      cellChksum := pCell^.udData + pCell^.udCRC32;
      IF ((pCell^.udCRC32 = 1954) & (pCell^.udType AND CELLMASK_VALID) & (cellChksum = pCell^.udChk)) THEN
        // in der 501.Zelle ist ein Zeiger auf den nächsten XRam-Block
        pHdr := sramStart + pCell^.udData;
        IF ((pHdr < sramStart) | (pHdr >= sramEnd)) THEN
          // Verkettung ungültig
      		sramErrorCode := EC_INV_BLK_CHAIN;
          SramError();
          AlarmSramError(pCell$DINT);
        END_IF;
      ELSE
        pHdr := NIL;
      END_IF;
    ELSE
      // Block war nur teilweise gefüllt, es handelt sich also um den letzten Block
      pHdr := NIL; // bewirkt Schleifenaabruch
    END_IF;

  END_WHILE;

END_FUNCTION

//------------------------------------------------------------------------------
// SramChecker
//------------------------------------------------------------------------------
FUNCTION GLOBAL SramCheckerCyclic
VAR
	pFileCell 	: ^XFileCell;
	pRamCell	: ^XRamCell;
	quit		: BOOL;
	chkSum		: UDINT;
	fileCellCnt	: UDINT;
END_VAR

	// wenn bereits ein Fehler festgestellt wurde, dann nichts mehr prüfen,
	// damit das Logfile nicht voll wird
	IF loaderRamexError <> 0 THEN
		AlarmSramError(1);	// Alarm immer wieder auslösen
		RETURN;
	END_IF;

 	IF _S_RAM_Hptr = NIL THEN
		RETURN;
	END_IF;

 	IF _S_RAM_Hptr^.DataValid < 2 THEN
    SramCheckV1();
		RETURN;
	END_IF;

 	IF !!isRamfileDatUsed THEN
		RETURN;
	END_IF;

	IF pRamFile^.udEntries = 0 THEN
		RETURN;
	END_IF;

(*
	pr, 7.2.05: ab 1.1.3 wird bei udEntries = 0 kein Sramfehler gemeldet
	IF _S_RAM_Hptr^.dataStart^.udEntries = 0 THEN
		sramErrorCode := 10;
		LogSramError();
		AlarmSramError(1);
		RETURN;
	END_IF;
*)

	IF (_S_RAM_Hptr^.dataStart^.udEntries XOR _S_RAM_Hptr^.dataStart^.udChk) <> 16#FFFFffff THEN
		sramErrorCode := EC_INV_BLK0_CHKSUM2;
		LogSramError();
		AlarmSramError(1);
		RETURN;
	END_IF;

	fileCellCnt := 0;
	quit := FALSE;
	WHILE !!quit DO

		pFileCell := #pRamFile^.aData[fileCellChkIdx];
		IF (pFileCell^.udCRC32 <> 0) & ((pFileCell^.udType AND 16#3C00_0000) = isXram) THEN
			// Ramex Zelle gefunden -> Checksumme prüfen, dann Schleife abbrechen
			pRamCell := _S_RAM_Hptr^.dataStart + pFileCell^.udpRelSram;

			chkSum := (pRamCell^.udType AND 16#00ffFFFF) + pRamCell^.udData + pRamCell^.udCRC32;
			IF chkSum <> pRamCell^.udChk THEN
				LogSramRamexError(pRamCell);
				AlarmSramError(pRamCell$DINT);
				//(0$^UDINT)^ := 0;	// Exception auslösen
			END_IF;

			quit := TRUE;
		END_IF;

		fileCellChkIdx += 1;
		IF fileCellChkIdx >= pRamFile^.udEntries THEN
			// das Ende ist erreicht -> index auf 0, dann Schleife abbrechen
			fileCellChkIdx := 0;
			quit := TRUE;
		END_IF;

		fileCellCnt += 1;
		IF fileCellCnt > 15 THEN
			// max. 15 File-Cells pro Durchlauf prüfen (sonst kann ein RUNTIME Error auftreten !)
			quit := TRUE;
		END_IF;

	END_WHILE;

END_FUNCTION
#endif

#ifdef _LSL_TARGETARCH_ARM
(*
  Überprüft den Inhalt der Sram-V2 Datenstruktur ob diese gültig ist
  und markiert den verwendeten Sram-Speicher in der MAT als belegt.

  Wenn der Sram Inhalt inhalt gültig ist, wird 0 zurückgegeben, sonst
  ein entsprechender Fehlercode.
*)
FUNCTION CHK_S_RAMV2
VAR_OUTPUT
  errCode : UDINT;
END_VAR
VAR
  i : UDINT;
  pXRAMHDR : ^XRAMHDR;
  pXRamCell : ^XRamCell;
  pXFileCell : ^XFileCell;
  ramStart :^XRamHdr;
END_VAR

  errCode := 0;

  IF !!(_S_RAM_Hptr^.DataValid AND 1) THEN
    errCode := EC_NOT_VALID;
    RETURN;
  END_IF;

  // In UsedData ist der Header mit eingerechnet
  IF _S_RAM_Hptr^.UsedData > _S_RAM_Hptr^.DataLength + _S_RAM_Hptr^.DataStart$UDINT - _S_RAM_Hptr$UDINT THEN
    errCode := EC_OUT_OF_SRAM;
    RETURN;
  END_IF;

  pXRAMHDR := _S_RAM_Hptr^.DataStart;
  IF pXRAMHDR^.udChk <> NOT pXRAMHDR^.udEntries THEN
    errCode := EC_INV_BLK0_CHKSUM;
    RETURN;
  END_IF;

  ramStart := _S_RAM_Hptr^.DataStart;

  // alle einträge o.k. jetzt machen wir noch eine Belegung im RAM mit dem mapper

  // *****************************************
  // die ersten 8 byte sind besonders //
  // *****************************************
  SRAM_MARKMemory(NIL, 8); //length: XRAMHDR (udEntries + udChk)

  pXFileCell := #pRamFile^.aData[0];
  FOR i := 1 TO pRamFile^.udEntries DO
    IF pXFileCell^.udCRC32 <> 0 THEN
      IF (pXFileCell^.udType AND 16#3C00_0000) <> ISXRAM THEN
        // normale RAMZelle	einfach speicher reservieren

        SRAM_MARKMemory(pXFileCell^.udpRelSram$^USINT, 4);

      ELSE
        // RAMEx Zelle

        pXRamCell := ramStart + pXFileCell^.udpRelSram;

        // 'XRamCell.udCRC32 = XFileCell.udCRC32' darf nicht geprueft werden weil
        // durch exchdataptr woanders liegen kann

        // CRC pruefen
        IF pXRamCell^.udChk = ((pXRamCell^.udType AND 16#00ffFFFF) +
                               pXRamCell^.udData +
                               pXRamCell^.udCRC32) THEN
          // super o.k. --> reservieren 16 byte block + reservieren Datenblock
          SRAM_MARKMemory(pXFileCell^.udpRelSram$^USINT, sizeof(XRamCell));
          SRAM_MARKMemory((pXRamCell^.udType AND 16#00FF_FFFF)$^USINT, pXRamCell^.udData AND 16#ffff);
        ELSE
          // die Ramex weist Fehler auf
          errCode := EC_INV_XRAMCELL_CHKSUM;
          LogSramRamexError(pXRamCell);

          pXFileCell^.udpRelSram := 0; // ungültig machen neuer speicher anlegen
          pXFileCell^.udCRC32 := 0; // loeschen damit nicht mehr gefunden wird

          pRamFile^.uiChange := 16#1234; // merker das Änderung

          pXRamCell^.udType := 0; // daten auch loaschen
          pXRamCell^.udData := 0; // daten auch loaschen
          pXRamCell^.udCRC32 := 0;
          pXRamCell^.udChk := 1;	 // damit chk sicher falsch ist
        END_IF;
      END_IF;
    END_IF;
    pXFileCell += sizeof(XFileCell);
  END_FOR;

END_FUNCTION

#ifdef _LSL_TARGETARCH_ARM_SUPPORTS_SRAMV1
(*
  Initialisiert das Sram im alten Format mit einem leeren Block.
*)
FUNCTION S_RAMV1_INITIALIZE_WITH_ONE_BLOCK
VAR
	sramSize : UDINT;
END_VAR

  _S_RAM_Hptr^.UsedData := 0;
  _S_RAM_Hptr^.DataValid := _S_RAM_Hptr^.DataValid AND 16#8000_0000; // alles außer Reorg-Flag rücksetzen

  IF _S_RAM_Hptr^.DataLength < maxSramSize THEN
    sramSize := _S_RAM_Hptr^.DataLength;
  ELSE
    sramSize := maxSramSize;
  END_IF;
  SRAM_STARTUP(sramSize, 1); // MAT für die Größe des SRAMs anlegen
  InitXramBlock();

END_FUNCTION
#endif // _LSL_TARGETARCH_ARM_SUPPORTS_SRAMV1

#ifdef _LSL_TARGETARCH_ARM_SUPPORTS_SRAMV1
(*
  Überprüft den Inhalt der Sram-V1 Datenstruktur ob diese gültig ist
  und markiert den verwendeten Sram-Speicher in der MAT als belegt.

  Wenn der Sram Inhalt inhalt gültig ist, wird 0 zurückgegeben, sonst
  ein entsprechender Fehlercode.
*)
FUNCTION CHK_S_RAMV1
VAR_OUTPUT
  errCode : UDINT;
END_VAR
VAR
  i : UDINT;
  pXRAMHDR : ^XRAMHDR;
  pXRamCell : ^XRamCell;
  cellValid : BOOL;
  typeFlags : UDINT;
  len : UDINT;
  ofs : UDINT;
END_VAR

  errCode := 0;

  IF !!(_S_RAM_Hptr^.DataValid AND 1) THEN
    errCode := EC_NOT_VALID;
    RETURN;
  END_IF;

  // In UsedData ist der Header mit eingerechnet
   IF _S_RAM_Hptr^.UsedData > _S_RAM_Hptr^.DataLength + _S_RAM_Hptr^.DataStart$UDINT - _S_RAM_Hptr$UDINT THEN
     errCode := EC_OUT_OF_SRAM;
     RETURN;
   END_IF;

  _S_RAM_Hptr^.DataStart^.aData[X_RAM_CELLS].udType :=
    _S_RAM_Hptr^.DataStart^.aData[X_RAM_CELLS].udType AND 16#80FFffff;  // 16*65535 Entries Total(used for quicksearch)

  //- Header prüfen --
  pXRAMHDR := _S_RAM_Hptr^.DataStart;
  WHILE 1 DO

    IF pXRAMHDR^.udEntries > X_RAM_CELLS THEN
      // more than 500 entries in one list !
      errCode := EC_INV_BLK_ENTRIES;
      RETURN;
    END_IF;
    IF pXRAMHDR^.udEntries <> NOT pXRAMHDR^.udChk THEN
      // CHKSUMME nicht OK
      errCode := EC_INV_BLK_CHKSUM;
      RETURN;
    END_IF;

    IF pXRAMHDR^.udEntries = 0 THEN
      S_RAMV1_INITIALIZE_WITH_ONE_BLOCK();	// #FA kommt vor weil active.dat nur header hat und ekien eintrage
      RETURN;
    END_IF;

    //-- Speicherblock belegen  mit länge eines blockes !
    SRAM_MARKMemory(pXRAMHDR$^USINT - _S_RAM_Hptr^.DataStart$UDINT, SIZEOF(XRAMHDR));

    pXRamCell := #pXRAMHDR^.aData[0];
    i := 0;
    WHILE i < pXRAMHDR^.udEntries DO
      cellValid := TRUE;
      IF (pXRamCell^.udType AND RamValid) = 0 THEN // ValidFlg (Bit 31) Must Be High !
        cellValid := FALSE;
      ELSIF pXRamCell^.udChk <> ((pXRamCell^.udType AND 16#00ffFFFF) +
                                 pXRamCell^.udData + pXRamCell^.udCRC32) THEN
        cellValid := FALSE;
      ELSE
        pXRamCell^.udType := pXRamCell^.udType AND NOT RAMUSED; // Clr Used Bit
        // CHK FOR Xtended Ram
        typeFlags := pXRamCell^.udType AND 16#3C00_0000;
        IF typeFlags <> 0 THEN
          IF typeFlags <> IsXram THEN
            cellValid := FALSE;
          END_IF;
        END_IF;
      END_IF;

      IF cellValid THEN
        len := pXRamCell^.udData AND 16#ffff; // mehr als 16#ffff geht nicht
        ofs := pXRamCell^.udType AND 16#00FF_ffff;
        SRAM_MARKMemory(ofs$^USINT, len);
      ELSE
        //--- contens of cell not valid , mark it as free (unused) --
        pXRamCell^.udType := 0;
        pXRamCell^.udData := 0;
        pXRamCell^.udCRC32 := 0;
        pXRamCell^.udChk := 0;
#ifdef SRAM_REPORT_INVALID_CELL1
        // Wenn ein Fehler bei einer Format-1 Zelle gefunden wird, dann wird standardmäßig
        // der Zelleninhalt auf 0 gesetzt und kein Sram Fehler gemeldet.
        // Warum wird kein Fehler gemeldet ?
        // Es hat einmal eine Loaderversion gegeben, bei der eine Sram-Zelle die noch nie
        // beschrieben wurde (also den Init-Wert aufweist), eine ungültige Chksum hatte.
        // Fürs Projekt hatte das keine neg. Auswirkungen, da die Chksum bereichtigt wurde,
        // sobald die Zelle beschrieben wurde (siehe Änderung in 02.02.102, SA17043).
        // Würde man jetzt bei einer falschen Chksum in einer Zelle einen Sram-Fehler melden
        // und das ganze Sram resettieren, dann könnte bei funktionierenden Applikationen
        // das Sram zurückgesetzt werden.
        errCode := EC_INV_V1_CELL;
        RETURN;
#endif
      END_IF;

      pXRamCell += sizeof(XRamCell);
      i += 1;
    END_WHILE;

    // -- CHK FOR NEXT BLOCK --
    IF i < X_RAM_CELLS THEN
      RETURN;
    END_IF;

    IF (pXRamCell^.udCRC32 <> 1954) | !!(pXRamCell^.udType AND RamValid) |
       (((pXRamCell^.udType AND 16#00ff_FFFF) + pXRamCell^.udData + pXRamCell^.udCRC32) <> pXRamCell^.udChk) THEN
      // Mark Cell 500 As EMPTY
      pXRamCell^.udType := 0;
      pXRamCell^.udData := 0;
      pXRamCell^.udCRC32 := 0;
      pXRamCell^.udChk := 0;
      RETURN;
    END_IF;

    pXRamCell := _S_RAM_Hptr^.DataStart + pXRamCell^.udData;

  END_WHILE;

END_FUNCTION
#endif // _LSL_TARGETARCH_ARM_SUPPORTS_SRAMV1
#endif

//-------------------------------------------
// Inhalt der daten im S-RAM -Prüfen und verwendeten Sram-Speicher in der MAT
// als belegt markieren.
//-------------------------------------------

//  udType:
//
// Bit 31.. 1= VALID  (CHksum is OK)
//     30.. 1= USED   (After Startup, it is conected to an Objekt)

//     29..   0   1    			(3000 0000)
//     28..   0   1
//     27..   0   0
//	   26..   0   0
//			  !   +-- 	RAMEX ; UdData field contains LENGTH of data,
//			  +--- RAM
//     25..   Frei
//	   24..   Frei
//
//	   0-23   Relative Startadress  of datablock if RAMEX

// CHK := udCrc+udData+(udType AND 16#00ffffff)

#ifdef _LSL_TARGETARCH_ARM
FUNCTION CHK_S_RAM
VAR_INPUT
  fDoNotReportErrors : UDINT;
END_VAR
VAR_OUTPUT
  wasValid : UDINT;
END_VAR
VAR
	sramSize : UDINT;
  errCode : UDINT;
END_VAR

  LogSramChk();
  wasValid := 1;
  sramErrorCode := 0;

  IF _S_RAM_Hptr^.DataLength < maxSramSize THEN
    sramSize := _S_RAM_Hptr^.DataLength;
  ELSE
    sramSize := maxSramSize;
  END_IF;
  SRAM_STARTUP(sramSize, 1); // MAT für die Größe des SRAMs anlegen

  IF isRamfileDatUsed & ((_S_RAM_Hptr^.DataValid SHR 16) AND 16#7fff) >= 2 THEN // Bit31 von DataValid ist das Reorg-Flag
    // =========================================================================
    // neue Version (mit ramfile.dat)
    // =========================================================================
    errCode := CHK_S_RAMV2();
    IF errCode <> 0 THEN
      sramErrorCode := errCode;
      wasValid := 0;

      IF errCode < 100 THEN
        IF !!fDoNotReportErrors THEN
          LogSramError();
        END_IF;
        // im file alles auf 0
        pRamFile^.udEntries := 0;
        pRamFile^.CRC32 := 0;
        pRamFile^.pLastEntry := 0;
        pRamFile^.uiChange := 16#1234; // merker das Änderung

        // auch im ram alles auf 0
        _S_RAM_Hptr^.UsedData := 0;
        _S_RAM_Hptr^.DataValid := (_S_RAM_Hptr^.DataValid AND 16#8000_0000) OR 16#0002_0000; // alles außer Reorg-Flag rücksetzen
      // und die anzahl der einträge auch loeschen
        _S_RAM_Hptr^.DataStart^.udEntries := 0;
        _S_RAM_Hptr^.DataStart^.udChk := 16#FFFF_ffff;

        IF _S_RAM_Hptr^.DataLength < maxSramSize THEN
          sramSize := _S_RAM_Hptr^.DataLength;
        ELSE
          sramSize := maxSramSize;
        END_IF;
        SRAM_STARTUP(sramSize, 1); // MAT für die Größe des SRAMs anlegen
        SRAM_MARKMemory(NIL, 8); //length: XRAMHDR (udEntries + udChk)
      END_IF;
    END_IF;

    // RAM allociert und als belegt gemeldet jetzt kommen die Konstruktoren der
    // RAM und RAMEX und wollen sich die Pointer holen
  ELSE
#ifdef _LSL_TARGETARCH_ARM_SUPPORTS_SRAMV1
    // =========================================================================
    // alte Version (ohne ramfile.dat)
    // =========================================================================
    errCode := CHK_S_RAMV1();
    IF errCode <> 0 THEN
      sramErrorCode := errCode;
      wasValid := 0;

      IF !!fDoNotReportErrors THEN
        LogSramError();
      END_IF;

      S_RAMV1_INITIALIZE_WITH_ONE_BLOCK();

    END_IF;
#else
    // altes Sram Format wird nicht unterstützt
    sramErrorCode := EC_UNSUPPORTED_FORMAT_V1;
    wasValid := 0;
    IF !!fDoNotReportErrors THEN
      LogSramError();
    END_IF;
#endif

  END_IF;

  GET_USED_S_RAM();

END_FUNCTION
#else
FUNCTION AWL CHK_S_RAM
VAR_INPUT
 fDoNotReportErrors : UDINT;
END_VAR
VAR_OUTPUT
 wasValid : UDINT;
END_VAR
VAR
 MAX_MEM	:UDINT ;
 RamStart   :^XramHdr;
END_VAR

		//*************************
		CALL		LogSramChk
		//*************************

		L.D			wasValid, 1

//	  SRAM_STARTUP(	16#40000 , 1);

		l.eax		_S_RAM_Hptr
		l.eax		(eax+MRAM_DESCR.DataLength)
		cmp.eax		maxSramSize
		jbe			CHK_S_RAMn
		l.eax		maxSramSize
CHK_S_RAMn
		PUSH		EAX			 // result
		PUSH.D		1
		PUSH.D		EAX 		 // Länge von OS
		CALL		SRAM_STARTUP
		ADD.ESP		2*4
		POP			EAX			 // RESULT

		L.D			MAX_MEM,0

   		L.EDI 		_S_RAM_Hptr
// test ob Ramfile.dat verwendet wird
		cmp.b		isRamfileDatUsed, 0
		je			chk_s_ram1

		l.ecx		(EDI+MRAM_DESCR.DataValid)
		shr.ecx		16
		cmp.ecx		2
		jb			chk_s_ram1			 // alte version

// es ist schon eine neue version
		l.ecx		(EDI+MRAM_DESCR.DataValid)
		and.ecx		1
		//*****
		L.D			sramErrorCode,EC_NOT_VALID
		//*****
		jz			chk_s_ram_error		// not valid

    (*DB1875*)
		l.eax		(EDI+MRAM_DESCR.DataLength)
		l.ecx		(EDI+MRAM_DESCR.UsedData)
    add.eax (EDI+MRAM_DESCR.DataStart)  // Header ist in UsedData mit eingerechnet
    sub.eax EDI
    cmp.ecx eax
		//*****
		L.D			sramErrorCode,5
		//*****
		jg			chk_s_ram_error

   		L.EDI		(EDI+MRAM_DESCR.DataStart)
		L.EAX		(EDI+XRAMHDR.udEntries)
		x.EAX		16#ffffffff
		cmp.EAX		(EDI+XRAMHDR.udChk)
		//*****
		L.D			sramErrorCode,EC_INV_BLK0_CHKSUM
		//*****
		jne			chk_s_ram_error

// alle einträge o.k. jetzt machen wir noch eine Belegung im RAM mit dem mapper
		L.EBX		pRamFile
		l.ECX		(EBX+XFILEHDR.udEntries)

		// pr, 21.1.06:
		//	Hier war eine Abfrage ob XFILEHDR.udEntries 0 ist und ein Jump
		//	auf chk_s_ram_error falls es 0 ist. Im Kommentar steht, daß das
		//  ein Fehler ist, der nicht sein kann.
		//	Wieso soll das ein Fehler sein ?
		//	Meiner Meinung nach ist das ganz normal daß XFILEHDR.udEntries 0 ist
		//  wenn ich ein Projekt ohne RAM- und RAMEX- Zellen habe.
		//	Ich war daher so frei und habe diese Abfrage einfach auskommentiert.
		//*****
		//L.D			sramErrorCode,4
		//*****
		//jecxz		chk_s_ram_error		// --> fehler der nicht sein kann

// *****************************************
// die ersten 8 byte sind besonders //
// *****************************************

		PUSH		EAX		// RESULT
		PUSH.D		8		// XRAMHDR: STRUCT =udEntries UDINT+udChk UDINT;
		CLR			EAX		// OFFSET 0 = 8 Byte
		PUSH		EAX
		CALL		SRAM_MARKMemory
		ADD.ESP		2*4
		POP			EAX		// Result

		ADD.EBX		XFILEHDR.aData		// EBX zeigt auf die ersten Dateneintrag

		O.ECX		ECX
		JZ			chk2lp_end
chk2lp
		l.eax		(ebx+XFileCell.udCRC32)		// CRC
		o.eax		eax							// flags setzen vergessen 01.10.2004 (aschl) damit geht eine Lawine los alles hin
		jz			chk2nxt				        // --> CRC = 0 invalid !! (nur zur Sicherheit)

		l.eax		(ebx+XFileCell.udType)		// finden ob RAM oder RAMEX
		A.EAX		16#3C00_0000
		cmp.eax		isXram						// test ob RAMEX
		je			chk2ramex					// --> ramEX

		l.eax		(ebx+XFileCell.udpRelSram)

// normale RAMZelle	einfach speicher reservieren
		PUSH		EAX							// RESULT
		PUSH.D		4							// XRAMHDR: STRUCT =udEntries UDINT+udChk UDINT;
		PUSH		EAX							// relativer RAMoffset
		CALL		SRAM_MARKMemory
		ADD.ESP		2*4
		POP			EAX							// Result
		jmp			chk2nxt

chk2ramex

		l.edi		_S_RAM_Hptr
		l.edi		(edi+MRAM_DESCR.DataStart)
		add.edi		(ebx+XFileCell.udpRelSram)  // EDI zeigt jetzt auf die Zelle

// jetzt zeigen wir in S_RAM da steht der Inhalt der gesamten Zelle

// darf nicht geprueft werden weil durch exchdataptr woanders liegen kann
//		l.eax		(edi+XRamCell.udCRC32)
//		cmp.eax		(ebx+XFileCell.udCRC32)
//		jne			chk2ramexFault				// CRC-RAM <> CRC-File

// CRC pruefen

		L.EAX		(EDI+XRamCell.udType)
		A.EAX		16#00ffFFFF
		ADD.EAX		(EDI+XRamCell.udData)
	   	ADD.EAX		(EDI+XRamCell.udCRC32)
		cmp.eax		(EDI+XRamCell.udChk)
		//*****
		L.D			sramErrorCode,EC_INV_XRAMCELL_CHKSUM
		//*****
		jne			chk2ramexFault				// checksumme falsch

// super o.k. --> reservieren 16 byte block + reservieren Datenblock

		PUSH		EAX		                 	// Result
		PUSH.D		sizeof (XRamCell)
		L.EAX		(EBX+XFileCell.udpRelSram)  // Startoffset Zelle
		PUSH		EAX
		CALL		SRAM_MARKMemory
		ADD.ESP		2*4
		POP			EAX							// Result

		PUSH		EAX		                 	// Result
		l.eax		(EDI+XRamCell.udData) 		// = LÄNGE
		and.eax		16#ffff                   	// mehr geht nicht
		PUSH		EAX
		L.EAX		(EDI+XRamCell.udType) 		// Startoffset
		A.EAX		16#00FF_FFFF
		PUSH		EAX
		CALL		SRAM_MARKMemory
		ADD.ESP		2*4
		POP			EAX							// Result
		jmp			chk2nxt

// die Ramex weist Fehler auf
chk2ramexFault
		//*************************
		PUSHAD
		PUSHFD
		PUSH		EDI
		CALL		LogSramRamexError
		POP			EDI
		POPFD
		POPAD
		//*************************
		L.D			wasValid, 0

		l.d			(ebx+XFileCell.udpRelSram),0 // ungültig machen neuer speicher anlegen
		l.d			(ebx+XFileCell.udCRC32),0	 // loeschen damit nicht mehr gefunden wird

		PUSH		EBX
		L.EBX		pRamFile
		L.W			(EBX+XFILEHDR.uiChange),16#1234		// merker das Änderung
		POP			EBX

		L.D			(EDI+XRamCell.udType) ,0	 // daten auch loaschen
		L.D			(EDI+XRamCell.udData) ,0
	   	L.D			(EDI+XRamCell.udCRC32),0
		L.D			(EDI+XRamCell.udChk)  ,1	 // damit chk sicher falsch ist

chk2nxt
		add.ebx		sizeof (XFileCell)
		loop		chk2lp
chk2lp_end
// RAM allociert und als belegt gemeldet jetzt kommen die Konstruktoren der
// RAM und RAMEX und wollen sich die Pointer holen
		JMP			S_RAM_CHK_RET

chk_s_ram_error
		L.EAX		fDoNotReportErrors
		O.EAX		EAX
		JNZ			Keine_Fehlermeldung_ins_Logfile
		//*************************
		PUSHAD
		PUSHFD
		CALL		LogSramError
		POPFD
		POPAD
		//*************************
Keine_Fehlermeldung_ins_Logfile

		L.D			wasValid, 0

// im file alles auf 0
		L.EDI		pRamFile
		l.d			(EDI+XFILEHDR.udEntries),0
		l.d			(EDI+XFILEHDR.CRC32),0
		l.d			(EDI+XFILEHDR.pLastEntry),0
		l.w			(EDI+XFILEHDR.uiChange),16#1234		// merker das Änderung

// auch im ram alles auf 0
   		L.EDI 		_S_RAM_Hptr
   		L.D			(EDI+MRAM_DESCR.UsedData),0
   		L.W			(EDI+MRAM_DESCR.DataValid+0),0
   		A.W			(EDI+MRAM_DESCR.DataValid+2),16#8000 // alles außer Reorg-Flag rücksetzen
   		O.W			(EDI+MRAM_DESCR.DataValid+2),2

// und die anzahl der einträge auch loeschen
		L.EDI		(EDI+MRAM_DESCR.DataStart)
		clr			eax
		s.eax		(EDI+XRAMHDR.udEntries)
		not			eax
		s.eax		(EDI+XRAMHDR.udChk)

		l.edi		_S_RAM_Hptr
		l.EAX		(edi+MRAM_DESCR.DataLength)
		cmp.eax		maxSramSize
		jbe			CHK_S_RAM2
		l.eax		maxSramSize

CHK_S_RAM2
		PUSH		EAX			// result
		PUSH.D		1
		PUSH.D		EAX         // max. SRAM Größe
		CALL		SRAM_STARTUP
		ADD.ESP		2*4
		POP			EAX			// RESULT

		PUSH		EAX		// RESULT
		PUSH.D		8		// XRAMHDR: STRUCT =udEntries UDINT+udChk UDINT;
		CLR			EAX		// OFFSET 0 = 8 Byte
		PUSH		EAX
		CALL		SRAM_MARKMemory
		ADD.ESP		2*4
		POP			EAX		// Result

		JMP			S_RAM_CHK_RET

CHK_S_RAM1

		l.ecx		(EDI+MRAM_DESCR.DataValid)
		and.ecx		1
		//*****
		L.D			sramErrorCode,EC_NOT_VALID
		//*****
		jz			S_RAM_INVALID		// not valid

    (*DB1875*)
		l.eax		(EDI+MRAM_DESCR.DataLength)
		l.ecx		(EDI+MRAM_DESCR.UsedData)
    add.eax (EDI+MRAM_DESCR.DataStart)  // Header ist in UsedData mit eingerechnet
    sub.eax EDI
    cmp.ecx eax
		//*****
		L.D			sramErrorCode,5
		//*****
		jg			S_RAM_INVALID

   		L.EDI		(EDI+MRAM_DESCR.DataStart)
		S.EDI		RamStart
		A.D			(EDI+XRAMHDR.aData[X_RAM_CELLS].udType),16#80FFffff  // 16*65535 Entries Total(used for quicksearch)

//- Header prüfen --

HDR_CHK_LP
		L.ECX		(EDI+XRAMHDR.udEntries)
		CMP.ECX		X_RAM_CELLS
		//*****
		L.D			sramErrorCode,EC_INV_BLK_ENTRIES
		//*****
		JA			S_RAM_INVALID		// more than 500 entries in one list !
		L.EAX		ECX
		NOT         EAX
		CMP.EAX		(EDI+XRAMHDR.udChk)	// CHKSUMME nicht OK
		//*****
		L.D			sramErrorCode,EC_INV_BLK_CHKSUM
		//*****
		JNE			S_RAM_INVALID
		jecxz		S_RAM_INITIALIZE_WITH_ONE_BLOCK	// #FA kommt vor weil active.dat nur header hat und ekien eintrage

//-- Speicherblock belegen  mit länge eines blockes !

		PUSH		EAX		// RESULT
		PUSH.D		SIZEOF(XRAMHDR)		// resu:=SRAM_MARKMEMORY(STartadr,LNG)
		L.EAX		EDI
		SUB.EAX		RamStart
		PUSH		EAX
		CALL		SRAM_MARKMemory
		ADD.ESP		2*4
		POP			EAX		// Result

		L.EDX		ECX

	   	L.EBX		XRAMHDR.aData[0]

S_CELL_CHK_LP
		L.EAX		(EDI+EBx+XRamCell.udType)			// ValidFlg Must Be High !
		O.EAX		EAX
		JNS			S_CELL_NOT_VALID					// Call not VALD (bit 31=0)

		A.EAX		16#00ffFFFF
		ADD.EAX		(EDI+EBX+XRamCell.udData)
	   	ADD.EAX		(EDI+EBX+XRamCell.udCRC32)
		CMP.EAX		(EDI+EBX+XRamCell.udChk)
		Jne			S_CELL_NOT_VALID

		A.D			(EDI+EBX+XRamCell.udType),NOT RamUsed  // Clr Used Bit

//    CHK FOR Xtended Ram //
		L.EAX		(EDI+EBX+XRamCell.udType)
		A.EAX		16#3C00_0000
		JZ			CHK_NEXT_CELL

		CMP.EAX		IsXram
		JNE			S_CELL_NOT_VALID

//        resu:=SRAM_MARKMEMORY(STartadr,LNG)

		PUSH		EAX		// RESULT

//     #FA vorsicht die length hat 2 teile byte0/1 ist die allocated length
//                                         byte2/3 ist die used length
//										   also ein mask ist wichtig

		l.eax		(EDI+EBX+XRamCell.udData) // = LÄNGE
		and.eax		16#ffff                   // mehr geht nicht
		PUSH		EAX
		L.EAX		(EDI+EBX+XRamCell.udType) // STartoffset
		A.EAX		16#00FF_ffff
		PUSH		EAX
		CALL		SRAM_MARKMemory
		ADD.ESP		2*4
		POP			EAX		// Result
		JMP			CHK_NEXT_CELL

//--- contens of cell not valid , mark it as free (unused) --

S_CELL_NOT_VALID

		L.D			(EDI+EBX+XRamCell.udType) ,0
		L.D			(EDI+EBX+XRamCell.udData) ,0
	   	L.D			(EDI+EBX+XRamCell.udCRC32),0
		L.D			(EDI+EBX+XRamCell.udChk)  ,0
#ifdef SRAM_REPORT_INVALID_CELL1
    // Wenn ein Fehler bei einer Format-1 Zelle gefunden wird, dann wird standardmäßig
    // der Zelleninhalt auf 0 gesetzt und kein Sram Fehler gemeldet.
    // Warum wird kein Fehler gemeldet ?
    // Es hat einmal eine Loaderversion gegeben, bei der eine Sram-Zelle die noch nie
    // beschrieben wurde (also den Init-Wert aufweist), eine ungültige Chksum hatte.
    // Fürs Projekt hatte das keine neg. Auswirkungen, da die Chksum bereichtigt wurde,
    // sobald die Zelle beschrieben wurde (siehe Änderung in 02.02.102, SA17043).
    // Würde man jetzt bei einer falschen Chksum in einer Zelle einen Sram-Fehler melden
    // und das ganze Sram resettieren, dann könnte bei funktionierenden Applikationen
    // das Sram zurückgesetzt werden.
    JMP     S_RAM_INVALID
#endif

// -- Next CELL

CHK_NEXT_CELL
		ADD.EBX  	SIZEOF(XRamCell)
		LOOP		S_CELL_CHK_LP

// -- CHK FOR NEXT BLOCK --

		CMP.EDX		X_RAM_CELLS				// entry nr must be X_RAM_CELLS
		JB			S_RAM_CHK_RET

	   	CMP.D		(EDI+EBX+XRamCell.udCRC32),1954
		JNE			NO_MORE_BLOCKS
	    L.EAX      	(EDI+EBX+XRamCell.udType)   // MUST BE VALID
		O.EAX		EAX
		JNS			NO_MORE_BLOCKS
		A.EAX		16#00ff_FFFF							// chk summ Must Be ok
		L.EAX		(EDI+EBX+XRamCell.udData)
	   	ADD.EAX		(EDI+EBX+XRamCell.udCRC32)
		CMP.EAX		(EDI+EBX+XRamCell.udChk)
		JNE			NO_MORE_BLOCKS

		L.EAX		(EDI+EBX+XRamCell.udData)
		L.EDI		RamStart
		ADD.EDI		EAX
		JMP			HDR_CHK_LP

// Mark Cell 500 As EMPTY

NO_MORE_BLOCKS
		L.D			(EDI+EBX+XRamCell.udType) ,0
		L.D			(EDI+EBX+XRamCell.udData) ,0
	   	L.D			(EDI+EBX+XRamCell.udCRC32),0
		L.D			(EDI+EBX+XRamCell.udChk)  ,0
		JMP			S_RAM_CHK_RET

//--------------------------------------------------
//-- S-RAM is Invalid ,initialise it with ONE BLOCK
//--------------------------------------------------

S_RAM_INVALID
		L.EAX		fDoNotReportErrors
		O.EAX		EAX
		JNZ			Keine_Fehlermeldung_ins_Logfile2
		//*************************
		PUSHAD
		PUSHFD
		CALL		LogSramError
		POPFD
		POPAD
		//*************************
Keine_Fehlermeldung_ins_Logfile2

		L.D			wasValid, 0

S_RAM_INITIALIZE_WITH_ONE_BLOCK
   		L.EDI 		_S_RAM_Hptr
   		L.D			(EDI+MRAM_DESCR.UsedData),0
   		L.W			(EDI+MRAM_DESCR.DataValid+0),0
   		A.W			(EDI+MRAM_DESCR.DataValid+2),16#8000 // alles außer Reorg-Flag rücksetzen

//	  SRAM_STARTUP(	16#40000 , 1);

		l.EAX		(edi+MRAM_DESCR.DataLength)
		cmp.eax		maxSramSize
		jbe			S_RAM_INVALID1
		l.eax		maxSramSize

S_RAM_INVALID1
		PUSH		EAX			// result
		PUSH.D		1
		PUSH		EAX  		// max. SRAM Größe
		CALL		SRAM_STARTUP
		ADD.ESP		2*4
		POP			EAX			// RESULT

//		 RelAdress:=InitXramBlock();

		PUSH		EAX
		CALL		InitXramBlock
		POP			EAX			// RESULTAT

//--- CHK IS Finished, Find Length of data --

S_RAM_CHK_RET
	    CALL		GET_USED_S_RAM
   		L.EDI 		_S_RAM_Hptr

END_FUNCTION
#endif

//-------------------------------------------------------------
// Whenever new S-RAM is alocatetd,S_Ram saver must be informed
//-------------------------------------------------------------

FUNCTION GLOBAL GET_USED_S_RAM
VAR
     usedLength : UDINT;
END_VAR

  IF !!hasSram THEN
    RETURN;
  END_IF;

  // Belegte Speichergrösse (bezogen auf speicherstart) abfragen
  usedLength := SRAM_GetLastAddr();
  // Größe des Headers dazuzählen
  usedLength := usedLength + _S_RAM_Hptr^.DataStart$UDINT - _S_RAM_Hptr$UDINT;

  // UsedData im _S_RAM_Hptr aktualisieren
  _S_RAM_Hptr^.UsedData := usedLength;

  // Wenn das SRAM Reorg aktiviert ist, dann wird das DataValid Flag
  // erst gesetzt, wenn alle RAM- und RAMEX- Zellen angelegt worden sind.
  IF !!fReorgSram | fSramInitCompleted THEN
    // Die unteren 16 Bit von DataValid auf den Wert 1 setzen
    _S_RAM_Hptr^.DataValid$UINT := 1;
    // Reorg-Flag (oberstes Bit von DataValid) rücksetzen
    _S_RAM_Hptr^.DataValid := _S_RAM_Hptr^.DataValid AND 0x7FFF_FFFF;
  END_IF;

END_FUNCTION

//-------------------------
// Calc CKSUM of RAMEX Hdr End MakeIt Valid
//-------------------------

#ifdef _LSL_TARGETARCH_ARM
FUNCTION GLOBAL MakeRamExChk
VAR_INPUT
  pXramCell : ^XramCell;
END_VAR
VAR
	udChk : UDINT;
END_VAR

  udChk := pXramCell^.udType AND 16#00ffFFFF;
  udChk += pXramCell^.udData;
  udChk += pXramCell^.udCRC32;

  pXramCell^.udChk := udChk;
  pXramCell^.udType := pXramCell^.udType OR (IsXram+RamValid+RamUsed);

END_FUNCTION
#else
FUNCTION GLOBAL AWL MakeRamExChk
VAR_INPUT
  pXramCell : ^XramCell;
END_VAR

  L.EDI     pXramCell
  L.EAX     (EDI+XRamCell.udType)
  L.EDX     EAX
  A.EAX     16#00ffFFFF
  ADD.EAX   (EDI+XRamCell.udData)
  ADD.EAX   (EDI+XRamCell.udCRC32)
  S.EAX     (EDI+XRamCell.udChk)
  O.EDX     (IsXram+RamValid+RamUsed)
  S.EDX     (EDI+XRamCell.udType)

END_FUNCTION
#endif

//-------------------------------
// Diese funktion erzeugt einen neuen ramblock mit 501 einträgen
// beim aufruf zeigt ein pointer auf die letzte zelle des akuellen blockes
// hier wird im feld "Data" die relative start_adresse des neuen blockes eingetregen
// als crc 32 steht  1954
// Die chk besteht wieder als summe von Data und CRC
//
//------------------------------

FUNCTION GLOBAL IniNewRamBlock
VAR_INPUT
  PtLastRamcell :^xRamCell;
END_VAR
VAR_OUTPUT
  Reladress :UDINT;
END_VAR

  RelAdress:=InitXramBlock();
  If Reladress <> 0 then
    PtLastRamcell^.udCRC32:=1954;
    PtLastRamcell^.udData$UDINT:=RelAdress$UDINT;
    PtLastRamcell^.udChk$UDINT:=PtLastRamcell^.udData$UDINT+PtLastRamcell^.udCRC32;
    PtLastRamcell^.udType:=PtLastRamcell^.udType or 16#80000000;      // valid
  END_IF;

END_FUNCTION

//-------------------------------------
// Initialise one block of Xram entries
//-------------------------------------
//  1. Ramdatenblock (hdr+501 eintrage) anfordern
//  2. nr Einträge auf 0 setzen
//  3. Alle blöcke mit 0 füllen
//
//
FUNCTION InitXramBlockEx
VAR_INPUT
  pGotMemory : ^BOOL;  // Da beim Returnwert 0 nicht unterschieden werden kann, ob
                       // der Offset 0 gemeint ist oder Out-Of-Memory, wird mit diesem
                       // Flag angezeigt, ob Speicher allokiert werden konnte.
END_VAR
VAR_OUTPUT
  xBlockOffset :UDINT ; // Offset of header
END_VAR

VAR
	I			  : DINT;
	PtxCell		  : ^XRamCell;
	ptxRamHead	  : ^XRAMHDR;
END_VAR

  xBlockOffset$^usint:=( SRAM_GetMemoryEx(sizeof(xRamHdr), pGotMemory));
  IF pGotMemory^ THEN
    ptxRamHead:= _S_RAM_Hptr^.DataStart+xBlockOffset;

    ptxRamHead^.udEntries:=0;
    ptxRamHead^.udChk:= 0;                     	// #FA damit kein compiler Fehler
    ptxRamHead^.udChk:= NOT ptxRamHead^.udChk; 	// value := not value (siehe doku)
    PtxCell:=#ptxRamHead^.aData[0];

    For i:= 0 to X_RAM_CELLS do
      PtxCell^.udChk:=0;
      PtxCell^.udCRC32:=0;
      PtxCell^.udData:=0;
      PtxCell^.udType:=16#0; 					// invalid
      PtxCell+=SIZEOF(XRamCell);
    end_for;
  END_IF;

END_FUNCTION

FUNCTION GLOBAL InitXramBlock
VAR_OUTPUT
  xBlockOffset :UDINT ; // Offset of header
END_VAR
VAR
	gotMemory : BOOL;
END_VAR

  xBlockOffset := InitXramBlockEx(#gotMemory);

END_FUNCTION

FUNCTION GLOBAL GetVersion_sRam
VAR_OUTPUT
	Version		: UDINT;
END_VAR

  IF !!hasSram THEN
    Version := 0;
  ELSE
    Version := (_S_RAM_Hptr^.DataValid SHR 16) AND 16#7FFF; // das oberste Bit (Reorg-Flag) ausblenden
  END_IF;

END_FUNCTION

#ifdef _LSL_TARGETARCH_ARM
// ---------------------------------------------------------------
// Funktion überprüft bei RAMex ob CRC im File = CRC im RAM
//
// Wenn die CRC im File nicht mit der CRC im RAM übereinstimmt,
// dann werden alle Einträge im File durchgegangen und über deren
// Verweis ins SRAM (udpRelSram) nachgeschaut, ob man eine Ramex-
// Zelle im SRAM mit der fraglichen CRC findet. Wenn eine gefunden
// wird, dann werden bei dem zu prüfenden und dem gefundenen Eintrag
// im File die Verweise ins SRAM (udpRelSram) ausgetauscht.
//
// Anm.pr:
// Das Aktualisieren der Verweises ins SRAM wird wegen EXCHANGE_DATA_PTR
// in der RamEx gemacht, wo die Daten von 2 Ramexobjekten vertauscht
// werden (füer IPR genützt)
// ---------------------------------------------------------------
FUNCTION CRC_extended
VAR_INPUT
  pXFileCell : ^XFileCell;
	pRamFile0	: ^XFILEHDR;
	_S_RAM_Hptr0 : ^MRAM_DESCR;
END_VAR
VAR_OUTPUT
  result : BOOL;
END_VAR
VAR
  pXRamCell : ^XRamCell;
  pXFileCellTemp : ^XFileCell;
  i : UDINT;
  udCRC32 : UDINT;
  oldUdpRelSram : UDINT;
  ramStart :^XRamHdr;
END_VAR

  result := FALSE;

  ramStart := _S_RAM_Hptr0^.DataStart;

  udCRC32 := pXFileCell^.udCRC32;
  pXRamCell := ramStart + pXFileCell^.udpRelSram;
  IF udCRC32 = pXramCell^.udCRC32 THEN
    result := TRUE;
    RETURN;
  END_IF;

  // CRC stimmt nicht überein -> Zellen im RAM nach der CRC durchsuchen
  // und wenn gefunden, die relative Ram-Adresse in der File-Zelle aktualisieren
  pXFileCellTemp := #pRamFile0^.aData[0];
  FOR i := 1 TO pRamFile0^.udEntries DO
    pXRamCell := ramStart + pXFileCellTemp^.udpRelSram;
    IF udCRC32 = pXramCell^.udCRC32 THEN
      // udpRelSram wird ausgetauscht
      oldUdpRelSram := pXFileCell^.udpRelSram;
      pXFileCell^.udpRelSram := pXFileCellTemp^.udpRelSram;
      pXFileCellTemp^.udpRelSram := oldUdpRelSram;
      result := TRUE;
      RETURN;
    END_IF;
    pXFileCellTemp += sizeof(XFileCell);
  END_FOR;

END_FUNCTION
#else
// ---------------------------------------------------------------
// funktion überprüft bei RAMex ob CRC im File = CRC im RAM
// ---------------------------------------------------------------
// --> ECX zeigt auf die Ramadresse(SRAM)
//     EAX = CRC
FUNCTION AWL CRC_extended
VAR
  oldUdpRelSram : UDINT;
END_VAR

		cmp.eax		(ecx+XRamCell.udCRC32)
		je			CRC_extend_ret // die CRC stimmt -> return

    // die CRC stimmt nicht -> File-Zellen durchgehen und über udpRelSram im Sram die Sram-Zelle mit der CRC suchen
		push		ebx
		push		edi

    l.ebx		(ebx+edi+XFileCell.udpRelSram)
    s.ebx   oldUdpRelSram // udpRelSram merken, damit man einen Austausch durchführen kann

		l.ecx		(EDI+XFILEHDR.udEntries)
		l.ebx		XFILEHDR.aData
Find_crcextend_loop
		l.edx		(edi+ebx+XFILECELL.udtype)
		and.edx		16#3C00_0000
		cmp.edx		isXram
		jne			find_crcextended_next

// now we found an extended RAM
// check if this ram has the right CRC

		l.EDX		_S_RAM_Hptr                 //++pr:Ich glaube hier sollte man besser nicht _S_RAM_Hptr verwenden,
                                        //     sondern den vom Aufrufer verwendeten Parameter _S_RAM_Hptr0 !
		L.EDX		(EDX+MRAM_DESCR.DataStart)
		ADD.EDX		(ebx+edi+XFileCell.udpRelSram)  // pointer to XramCell

		cmp.eax		(EDX+XRamCell.udCRC32)
		jne			find_crcextended_next			// --> crc is different

// wir haben das richtige gefunden
		l.ecx		edx
    // werte in updRelSram austauschen
		l.eax		(ebx+edi+XFileCell.udpRelSram)
    l.edx   oldUdpRelSram
    s.edx		(ebx+edi+XFileCell.udpRelSram)

		pop			edi
		pop			ebx
		s.eax		(ebx+edi+XFileCell.udpRelSram)  // store the real pointer
		clc
		jmp			CRC_extend_end

find_crcextended_next
		add.ebx		sizeof (XFileCell)
		loop		Find_crcextend_loop				// weitersuchen
		pop			edi
		pop			ebx
		stc
		jmp			CRC_extend_end

CRC_extend_ret
		clc
CRC_extend_end
END_FUNCTION
#endif

//------------------------------------------------------------------------------
// Allokiert eine Ramzelle (für SRAM Version 2 = SRAM + FILE)
//	a) RAM
//		Im SRAM werden 4 Bytes belegt,
//		Im FILE werden 12 Bytes belegt
//	b) RAMEX
//		Im SRAM werden 16 Bytes belegt,
//		Im FILE werden 12 Bytes belegt
// Die Zelle im FILE (XRamCell) enthält die Offset-Adresse der Zelle im SRAM.
// Das Flag uiChange des File-Headers wird auf 16#1234 gesetzt, um anzuzeigen,
// das der File-Cache (pRamFile) aufs File geschrieben werden muß.
//
// Der SRAM Speicher für die RAMEX Daten wird hier nicht allokiert, dafür ist
// der Aufrufer zuständig.
//------------------------------------------------------------------------------
FUNCTION Add_sRamFile_I
VAR_INPUT
	CRC32		:  UDINT;
	ppRamAdr	: ^UDINT;
	ppFileAdr	: ^pXFileCell_t;
	uiType		: UDINT;				// 0=RamZelle 1=RamExZelle
END_VAR
VAR_OUTPUT
	state		: UDINT;
END_VAR
VAR
	nAlloc : UDINT;
  pRam : ^USINT;
  pXFileCell : ^XFileCell;
  pXRamCell : ^XRamCell;
  allocSize : UDINT;
END_VAR

  state := 0; // auf o.k.

  IF uiType = 0 THEN
    nAlloc := 4;
  ELSE
    nAlloc := 16;
  END_IF;

  IF pRamFile^.udEntries < X_FILE_CELLS_2 THEN
    IF pRamFile^.udEntries = X_FILE_CELLS & LDR_allocated_XFileCells = X_FILE_CELLS THEN
      allocSize := XFILEHDR.adata + X_FILE_CELLS_2 * SIZEOF(XFileCell);
    	pRamFile := _realloc_LDR(pRamFile, allocSize)$^XFILEHDR;
      IF pRamFile <> NIL THEN
        LDR_allocated_XFileCells := X_FILE_CELLS_2;
        LDR_allocated_XFileSize := allocSize;
      END_IF;
    END_IF;
    pRam := SRAM_GetMemory(nAlloc);
  ELSE
    TRACE_ERR("Too many RAM objects");
    pRam := NIL;
  END_IF;
  IF pRam = 0 THEN
    ppRamAdr^ := NIL; // kein memory pointer
    ppFileAdr^ := NIL; // kein memory pointer
    state := 16#FFFFffff; // auf fehler stellen
    LDR_outOfSramMem := 1; // im Flag merken, dass keine Sram-Speicher mehr vorhanden ist
    RETURN;
  END_IF;

  pXFileCell := #pRamFile^.aData[pRamFile^.udEntries];

  //pr:
  //  Hier müsste GET_USED_S_RAM aufgerufen werden, weil SRAM_GetMemory
  //  etwas allokiert hat. Aus Performancegründen wird dieser Aufruf aber
  //  in die Funktion LDR_FreeSramKopie ausgelagert. Diese Funktion wird
  //  am Ende der SRAM Initialisierung aufgerufen.

  // merken im File
  pXFileCell^.udpRelSram := pRam$UDINT;

  _S_RAM_Hptr^.DataStart^.udEntries += 1;
  _S_RAM_Hptr^.DataStart^.udChk := NOT _S_RAM_Hptr^.DataStart^.udEntries;

  // jetzt absolut pointer berechnen
  pXRamCell := _S_RAM_Hptr^.DataStart + pRam$UDINT;
  ppRamAdr^ := pXRamCell$UDINT; // rückgabewert

  // wenn wir 16 byte haben muessen wir jetzt auch die CRC eintragen und alles andere loeschen
  IF uiType <> 0 THEN
		// wir reservieren 16 byte und tun so
		// als wäre das eine alte XramCell damit ist RamEx fast kompatibel
    pXRamCell^.udCRC32 := CRC32;
    pXRamCell^.udType := 0;
    pXRamCell^.udData := 0;
    pXRamCell^.udChk := 0;

    pXFileCell^.udType := ISXRAM;
  ELSE
    pXFileCell^.udType := 0;
  END_IF;
  pXFileCell^.udCRC32 := CRC32;

  ppFileAdr^ := pXFileCell; // rückgabewert

  pRamFile^.udEntries += 1; // eintrag erhöhen am ende
  pRamFile^.uiChange := 16#1234;	// merker das Änderung

END_FUNCTION

// ---------------------------------------------------------------------
//  suchen der eines Eintrages im File und daraus die Pointer ableiten
// ---------------------------------------------------------------------
//
//  Achtung bei uiType = 1 kann wenn die Ramex ein IPR Programm ist
//  durch exchange dataptr in der Ramex es passiren das die Ramex
//  jetzt woanders ist um somit der offset nicht mehr stimmt !!
//  Dann wird muessen alle Ramex durchsucht werden um herauszufinden
//  wo der neue steckt !!
//
#ifdef _LSL_TARGETARCH_ARM
FUNCTION Find_sRamFile_I
VAR_INPUT
	pRamFile0	: ^XFILEHDR;
	_S_RAM_Hptr0: ^MRAM_DESCR;
	CRC32		:  UDINT;
	ppRamAdr	: ^UDINT;
	ppFileAdr	: ^pXFileCell_t;
	uiType		: UDINT;				// 0=RamZelle 1=RamExZelle
END_VAR
VAR_OUTPUT
	state		: UDINT;
END_VAR
VAR
	nLoops : UDINT;
  pXFileCell : ^XFileCell;
  pLastEntry : UDINT;
END_VAR

  state := 0; // auf o.k.

  IF (pRamFile0^.pLastEntry > 0) & (pRamFile0^.pLastEntry < pRamFile0^.udEntries) THEN
    // wir haben uns den letzten stand der dinge vom suchen gemerkt und um
    // schneller zu sein suchen wir ab hier und dann erst vom beginn
    // ist bei vielen ramzellen 10.000 mal schneller
    nLoops := 2;
  ELSE
    // suchen von vorne
    pRamFile0^.pLastEntry := 0;
    nLoops := 1;
  END_IF;

  WHILE nLoops > 0 DO

    pLastEntry := pRamFile0^.pLastEntry;
    pXFileCell := #pRamFile0^.aData[pLastEntry];
    WHILE pLastEntry < pRamFile0^.udEntries DO
      pLastEntry += 1;

      IF (pXFileCell^.udCRC32 = CRC32) & ((uiType = 0) | (CRC_extended(pXFileCell, pRamFile0, _S_RAM_Hptr0))) THEN
        // gefunden jetzt geben wir die pointer zurück
        ppRamAdr^$UDINT := _S_RAM_Hptr0^.DataStart$UDINT + pXFileCell^.udpRelSram;
        ppFileAdr^ := pXFileCell;

        pRamFile0^.pLastEntry := pLastEntry;
        RETURN;
      END_IF;

      pXFileCell += sizeof(XFileCell);
    END_WHILE;

    // Zweiter Schleifendurchlauf von vorne
    pRamFile0^.pLastEntry := 0;
    nLoops -= 1;

  END_WHILE;

  // **************************************** //
  // nicht vorhanden --> neuen erfinden       //
  // **************************************** //

	state := 16#FFFFFFFE;			// auf nicht gefunden stellen

END_FUNCTION
#else
FUNCTION AWL Find_sRamFile_I
VAR_INPUT
	pRamFile0	: ^XFILEHDR;
	_S_RAM_Hptr0: ^MRAM_DESCR;
	CRC32		:  UDINT;
	ppRamAdr	: ^UDINT;
	ppFileAdr	: ^pXFileCell_t;
	uiType		: UDINT;				// 0=RamZelle 1=RamExZelle
END_VAR
VAR_OUTPUT
	state		: UDINT;
END_VAR

		l.d			state,0						// auf o.k.

		push		esi
		l.edi		pRamFile0
		l.ecx		(EDI+XFILEHDR.udEntries)
		jecxz		Find_sRamFile_add			// --> neues eintragen

// wir haben uns den letzten stand der dinge vom suchen gemerkt und um
// schneller zu sein suchen wir ab hier und dann erst vom beginn
// ist bei vielen ramzellen 10.000 mal schneller

		cmp.d		(edi+XFILEHDR.pLastEntry),0
		je			find_sRamFile_start0		// --> wir fangen bei 0 an
		sub.ecx		(edi+XFILEHDR.pLastEntry)
		js			find_sRamFile_start0		// --> von vorne suchen
		jecxz		find_sRamFile_start0		// --> von vorne suchen

		l.ebx		(edi+XFILEHDR.pLastEntry)
		l.eax		sizeof (XFileCell)
		mul			ebx
		l.ebx		eax
		add.ebx		XFILEHDR.aData
		l.eax		CRC32

Find_sRamFile_loop0
		cmp.eax		(ebx+edi+XFileCell.udCRC32)
		jne			Find_sRamFileNext0

		inc.d		(edi+XFILEHDR.pLastEntry)		// einer weiter vor

// gefunden jetzt geben wir die pointer zurück

		l.ecx		_S_RAM_Hptr0
		L.ECX		(ECX+MRAM_DESCR.DataStart)
		ADD.ECX		(ebx+edi+XFileCell.udpRelSram)

// falls type = 1 check ob auch CRC übereinstimmt
		cmp.d		uiType,0
		je			find_sramStd
		call		CRC_extended		     // pruefen ob wirklich der richtige
		jc			find_sRamFile_start0
find_sramStd
		l.EAX		ppRamAdr
		s.ECX		(EAX)

		l.eax		ppFileAdr
		add.ebx		edi
		s.ebx		(eax)

		jmp			Find_sRamFile_ret

Find_sRamFileNext0
		add.ebx		sizeof (XFileCell)
		// merken wo wir waren
		inc.d		(edi+XFILEHDR.pLastEntry)
		loop		Find_sRamFile_loop0

// hier starten wir ganz von vorne und durchsuchen alles

find_sRamFile_start0
		l.ecx		(EDI+XFILEHDR.udEntries)
		clr			edx
		l.ebx		XFILEHDR.aData
		l.eax		CRC32
Find_sRamFile_loop
		cmp.eax		(ebx+edi+XFileCell.udCRC32)
		jne			Find_sRamFileNext
// merken wo wir waren
		s.edx		(edi+XFILEHDR.pLastEntry)

// gefunden jetzt geben wir die pointer zurück

		l.ecx		_S_RAM_Hptr0
		L.ECX		(ECX+MRAM_DESCR.DataStart)
		ADD.ECX		(ebx+edi+XFileCell.udpRelSram)

// falls type = 1 check ob auch CRC übereinstimmt
		cmp.d		uiType,0
		je			find_sramStdB
		call		CRC_extended		     // pruefen ob wirklich der richtige
		jc			Find_sRamFile_add
find_sramStdB

		l.EAX		ppRamAdr
		s.ECX		(EAX)

		l.eax		ppFileAdr
		add.ebx		edi
		s.ebx		(eax)

		jmp			Find_sRamFile_ret

Find_sRamFileNext
		add.ebx		sizeof (XFileCell)
		inc			edx
		loop		Find_sRamFile_loop

// **************************************** //
// nicht vorhanden --> neuen erfinden       //
// **************************************** //

Find_sRamFile_add
		l.d			state,16#FFFFFFFE			// auf nicht gefunden stellen
		jmp			Find_sRamFile_ret

Find_sRamFile_ret
		pop			esi
END_FUNCTION
#endif

#ifdef LDR_RETSVR
(* Rundet einen Wert auf den nächsten 2^x Wert auf (z.B. 100 auf 128, 200 auf 256) *)
FUNCTION RoundUpPow2
VAR_INPUT
	value	: UDINT;
END_VAR
VAR_OUTPUT
	result : UDINT;
END_VAR

  result := 1;
  WHILE value > 0 DO
    value := value SHR 1;
    result := result SHL 1;
  END_WHILE;

END_FUNCTION

FUNCTION Add_File_I
VAR_INPUT
	CRC32		:  UDINT;
	ppRamAdr	: ^void;
END_VAR
VAR_OUTPUT
	state		: UDINT;
END_VAR
var
  Cell : XRamCell;
end_var

  state := 2; // hat nicht funktioniert!

  // Zelle vorbereiten
  Cell.udChk := 0;
  Cell.udCRC32 := CRC32;
  Cell.udData := 0;
  Cell.udType := _S_RAM_Hptr_File^.UsedData;  // im udType wird die Fileposition gespeichert!

  // Fileimage updaten

  _S_RAM_Hptr_File^.UsedData += sizeof( XRamCell );
  _S_RAM_Hptr_File := ReAlloc_S_RAM_Hptr_File(_S_RAM_Hptr_File, _S_RAM_Hptr_File^.UsedData);
  if( _S_RAM_Hptr_File = NIL )then
    return;
  end_if;
  _memcpy( _S_RAM_Hptr_File + Cell.udType, #Cell, sizeof( XRamCell ) );

  // Reorg. Image updaten

  _S_RAM_Hptr_File_New := ReAlloc_S_RAM_Hptr_File(_S_RAM_Hptr_File_New, _S_RAM_Hptr_File_New^.UsedData + sizeof( XRamCell ));
  if( _S_RAM_Hptr_File_New = NIL )then
    return;
  end_if;
  Cell.udType := _S_RAM_Hptr_File_New^.UsedData;
  _memcpy( _S_RAM_Hptr_File_New + _S_RAM_Hptr_File_New^.UsedData, #Cell, sizeof( XRamCell ) );
  _S_RAM_Hptr_File_New^.UsedData += sizeof( XRamCell );

  // Rückgabe
  _memcpy( ppRamAdr, #Cell, sizeof( XRamCell ) );
  state := 1;

END_FUNCTION

VAR_PRIVATE
  lastFindFileIndex : UDINT;
END_VAR

FUNCTION Find_File_I
VAR_INPUT
  pMem    : ^MRAM_DESCR;
	CRC32		:  UDINT;
	ppRamAdr	: ^void;
  bDontAdd   : BOOL;
END_VAR
VAR_OUTPUT
	state		: UDINT;
END_VAR
var
  pCell   : ^XRamCell;
  nCells : udint;
  i :  udint;
end_var

  // Die Suche wird nicht bei Index 0 sondern bei Index lastFindFileIndex gestartet.
  // lastFindFileIndex steht auf dem Wert vom letzten Aufruf dieser Funktion.
  // Dadurch wird die Suche beschleunigt, weil die Zellen normalerweise in der Reihenfolge
  // abgefragt werden, wie sie im Speicher angeordnet sind.
  ppRamAdr^ := NIL;
  state := 1;
  nCells := (pMem^.UsedData - pMem^.DataStart$udint) / sizeof( XRamCell );
  pCell := pMem + pMem^.DataStart$udint + lastFindFileIndex * sizeof( XRamCell );

  for i := 1 to nCells do
    if lastFindFileIndex >= nCells then
      lastFindFileIndex := 0;
      pCell := pMem + pMem^.DataStart$udint;
    end_if;

    // Zelle gefunden -> ins Reorg. eintragen und den richtigen Pointer zurückgeben
    if( pCell^.udCRC32 = CRC32 )then

      if !!bDontAdd then
        _S_RAM_Hptr_File_New := ReAlloc_S_RAM_Hptr_File(_S_RAM_Hptr_File_New, _S_RAM_Hptr_File_New^.UsedData + sizeof( XRamCell ));
        if( _S_RAM_Hptr_File_New = NIL )then
          return;
        end_if;
        pCell^.udType := _S_RAM_Hptr_File_New^.UsedData;  //den udType brauch ich hier nicht, da kommt der Offset im File rein!

        //Reorg.
        _memcpy( _S_RAM_Hptr_File_New + _S_RAM_Hptr_File_New^.UsedData, pCell, sizeof( XRamCell ) );

        // Datenlänge im Reorg. korrigieren
        _S_RAM_Hptr_File_New^.UsedData += sizeof( XRamCell );
      end_if;

      // Rückgabe
      _memcpy( ppRamAdr, pCell, sizeof( XRamCell ) );

      state := 0;
      exit;

    end_if;

    // nächster Eintrag
    lastFindFileIndex += 1;
    pCell += sizeof( XRamCell );

  end_for;

END_FUNCTION

// sucht einen remanenten Server im File
FUNCTION GLOBAL Find_FileEx
VAR_INPUT
	CRC32		:  UDINT;
	ppRamAdr	: ^void;
  bDontAdd   : BOOL;
END_VAR
VAR_OUTPUT
	state		: UDINT;
END_VAR
var
 	errCode : DINT;
	rc : DINT;
end_var

  // gibts den Handle überhaupt schon?
  if( hLDR_remSvr = NIL )then

    // wenn nicht muss das File zuerst initialisiert werden
    if( InitRetainSvrFile( 0 ) <> 1 )then
      state := 3;
      return;
    end_if;
  end_if;

  // Einlesen der remanenten Server und vorbereiten des Reorg.
  rc := LoadSramKopie( #errCode, hLDR_remSvr, 0 );
  if( rc <> 0 )then
    DEBUGLOG2( "%010d Retentive server file I/O error, rc=%d, errCode = 0x%X", rc$UDINT, errCode$udint );
  end_if;

  // suchen eines bestimmten Servers im File
  state := Find_File_I( _S_RAM_Hptr_File, CRC32, ppRamAdr, bDontAdd );

  if(bDontAdd = 0) then
  	if( state <> 0 ) then
  		// nicht gefunden, neue Zelle anlegen
  		nbrOfCells_notFound += 1;
	  	state := Add_File_I( CRC32, ppRamAdr );
  	end_if;
  end_if;

END_FUNCTION

FUNCTION GLOBAL Find_File
VAR_INPUT
	CRC32		:  UDINT;
	ppRamAdr	: ^void;
END_VAR
VAR_OUTPUT
	state		: UDINT;
END_VAR

  state := Find_FileEx(CRC32, ppRamAdr, FALSE);

END_FUNCTION

#endif //LDR_RETSVR

FUNCTION GLOBAL Find_sRamFileEx
VAR_INPUT
	CRC32		:  UDINT;
	ppRamAdr	: ^UDINT;
	ppFileAdr	: ^pXFileCell_t;
	uiType		: UDINT;				// 0=RamZelle 1=RamExZelle
  bDontAdd  : BOOL;
END_VAR
VAR_OUTPUT
	state		: UDINT;
END_VAR
VAR
	pRamAdr_Kopie	: ^XRamCell;
	pFileAdr_Kopie	: ^XFileCell;
	// Die folgenden beiden Variablen werden benötigt, weil die beiden Übergabeparameter
	// ppRamAdr und ppFileAdr nicht als Zeiger auf Zeiger deklariert wurden.
	// Wenn man die Werte auf die beide lokalen Variablen kopiert, dann kann man ohne
	// umständliche casterei damit arbeiten.
	pRamAddr	: ^XRamCell;
	pFileAdr : ^XFileCell;

	udAllocated : UDINT;
	udLength : UDINT;
	RelAdress		: UDINT;
	pData : ^USINT;
	pData_Kopie : ^USINT;
	errCode : DINT;
	rc : DINT;
    ret_sRamHptr : UDINT;
END_VAR

  // Diese Funktion wird für die RamEx Klasse benötigt und um den Loader kompatibel zu halten
  // 1 bewirkt, dass die Funktion "Find_sRamFileEx" beim Rückgabewert nicht 0 für gefunden liefert,
  // sonder entweder _s_Ram_hptr oder _s_Ram_hptr_Kopie (REORG) um auf die SRAM Daten zugreifen zu können.
  ret_SramHptr := 0;
  if((ppRamAdr <> NIL) & (ppRamAdr^ = 1)) then
    ret_SramHptr := 1;
  end_if;

	IF fReorgSram THEN
		rc := LoadSramKopie(#errCode, 0, 0);
		IF rc <> 0 THEN
			// das Laden de SRAM Kopie hat nicht funktioniert
			fReorgSram := 0;
			DEBUGLOG2("%010d LoadSramKopie failed, rc=%d, errCode = 0x%X" , rc$UDINT, errCode$UDINT);
		END_IF;
	END_IF;

	IF fReorgSram THEN
		// in der Kopie suchen
		state := Find_sRamFile_I(pRamFile_Kopie, _s_Ram_hptr_Kopie, CRC32, ppRamAdr, ppFileAdr, uiType);
	ELSE
		// im SRAM suchen
		state := Find_sRamFile_I(pRamFile, _s_Ram_hptr, CRC32, ppRamAdr, ppFileAdr, uiType);
	END_IF;

	if((state = 0) & (bDontAdd = TRUE)) then
    if(ret_sRamHptr = 1) then
    	if(fReorgSram) then
        state := _s_Ram_hptr_Kopie$UDINT;
      else
        state := _s_Ram_hptr$UDINT;
      end_if;
    end_if;

		return;
	end_if;

	IF state <> 0 | ppRamAdr^ = NIL THEN
		// nicht gefunden (weder im SRAM noch in der Kopie), neue Zelle anlegen
		nbrOfCells_notFound += 1;

    if(bDontAdd = FALSE) then
  		state := Add_sRamFile_I(CRC32, ppRamAdr, ppFileAdr, uiType);
    end_if;
	ELSIF fReorgSram THEN
		// in der Kopie gefunden, Zelle aus der Kopie ins SRAM kopieren
		nbrOfCells_foundInCopy += 1;

		pRamAdr_Kopie := ppRamAdr^$^XRamCell;
		pFileAdr_Kopie := ppFileAdr^;
		ppRamAdr^$^UDINT := NIL;
		ppFileAdr^$^XFileCell := NIL;

    if(bDontAdd = FALSE) then
  		state := Add_sRamFile_I(CRC32, ppRamAdr, ppFileAdr, uiType);
    end_if;
		pRamAddr := ppRamAdr^$^XRamCell;
		pFileAdr := ppFileAdr^$^XFileCell;

		IF state = 0 & pRamAddr <> NIL THEN
			IF uiType = 0 THEN
				// RAM
			    pRamAddr^$dint  :=pRamAdr_Kopie^$dint;
			    pFileAdr^.udType:=16#C0000000;    // ganz am ende machen wir uns gültig !
			ELSE
				// RAMEX
 		     	udLength := pRamAdr_Kopie^.udData shr 16;
				// wenn die Länge der Daten > 0 ist, dann muss das RAMEX Objekt mit
				// den Daten aus der Kopie vorgeladen und für gültig erklärt werden
				IF udLength > 0 THEN
				 	RelAdress$UDINT:= (SRAM_GetMemory(udLength))$UDINT;
				 	// --- Speicher ist zugewiesen worden --
				 	If RelAdress <> 0 THEN
				   		GET_USED_S_RAM();
				   		udAllocated		      := SRAM_GET_ALLOCATED(udLength);
			  	   		pRAMaddr^.udData$UDINT := (udLength shl 16) or (udAllocated and 16#ffff);
				   		pRAMaddr^.udType 	  := RelAdress;
				   		pData				  := _S_RAM_Hptr^.DataStart+RelAdress;
				   		pData_Kopie			  := _S_RAM_Hptr_Kopie^.DataStart+(pRamAdr_Kopie^.udType and 16#00FF_ffff);
				   		_memcpy(pData, pData_Kopie, udLength);   // Speicher aus dem Inhalt aus der Kopie vorladen
		           		MakeRamExChk(pRAMaddr);

				 	// -- Kein speicher verfügbar !!
				 	ELSE

	               		state := 0xFFFFFFFF;
			       		ppRamAdr^$^UDINT := NIL;
			       		ppFileAdr^$^XFileCell := NIL;

				 	END_IF;
				ELSE
	           		MakeRamExChk(pRAMaddr);
				END_IF;
			END_IF;
		END_IF;
	ELSE
		nbrOfCells_foundInSram += 1;
	END_IF;

END_FUNCTION

FUNCTION GLOBAL Find_sRamFile
VAR_INPUT
	CRC32		:  UDINT;
	ppRamAdr	: ^UDINT;
	ppFileAdr	: ^pXFileCell_t;
	uiType		: UDINT;				// 0=RamZelle 1=RamExZelle
END_VAR
VAR_OUTPUT
	state		: UDINT;
END_VAR

  state := Find_sRamFileEx(CRC32, ppRamAdr, ppFileAdr, uiType, FALSE);

END_FUNCTION

//------------------------------------------------------------------------------
// Allokiert eine Ramzelle (für SRAM Version 1 = SRAM ohne FILE)
//  Im SRAM werden 16 Bytes belegt
//
// Der SRAM Speicher für die RAMEX Daten wird hier nicht allokiert, dafür ist
// der Aufrufer zuständig.
//------------------------------------------------------------------------------
#ifdef _LSL_TARGETARCH_ARM
FUNCTION Add_sRam_I
VAR_INPUT
#pragma warning(disable:73)
	CRC32		: UDINT;
#pragma warning(default:73)
END_VAR
VAR_OUTPUT
	pRamAdr		: ^XramCell;
END_VAR
#ifdef _LSL_TARGETARCH_ARM_SUPPORTS_SRAMV1
VAR
   RamStart     : ^XramHdr;
   pXramHdr     : ^XRAMHDR;
   RelAdress	  :  UDINT;
END_VAR

  pRamAdr := 0$^XRamCell;
  RamStart := _S_RAM_Hptr^.DataStart;

  // Die folgende Schleife geht die Verkettung der XRAM-Blöcke durch
  // bis das Ende erreicht ist.
  pXramHdr := RamStart;
  WHILE 1 DO
		// Abbruch, wenn ein XRAM-Block weniger als 500 XRAM-Zellen enthält
		// oder wenn kein Zeiger auf einen weiteren XRAM-Block existiert.
    IF (pXramHdr^.udEntries < X_RAM_CELLS) | (pXramHdr^.aData[X_RAM_CELLS].udCRC32 <> 1954) THEN
      EXIT;
    END_IF;
    pXramHdr := RamStart + pXramHdr^.aData[X_RAM_CELLS].udData; // offset zum nächsten block
  END_WHILE;

// There is Place in our list, Write It

  IF pXramHdr^.udEntries = X_RAM_CELLS THEN
    // Neuen Block anlegen  und eintragen
    RelAdress := IniNewRamBlock(#pXramHdr^.aData[X_RAM_CELLS]);
    IF RelAdress = 0 THEN
      // out of memory !!!
      LDR_outOfSramMem := 1;    // im Flag merken, dass keine Sram-Speicher mehr vorhanden ist
      RETURN;
    END_IF;
    GET_USED_S_RAM();	// Memory updaten
    pXramHdr := RamStart + RelAdress;
  END_IF;

  pRamAdr := #pXramHdr^.aData[pXramHdr^.udEntries];

//------------------------------------------------------
// Block belegen und auf ungültig setzen
//------------------------------------------------------

  pRamAdr^.udCRC32 := CRC32;
  pRamAdr^.udData := 0;
  pRamAdr^.udChk := CRC32;
  pRamAdr^.udType := 0; // Type = RAM,Daten nicht gültig

  pXramHdr^.udEntries += 1;
  pXramHdr^.udChk := NOT pXramHdr^.udEntries;
#else // _LSL_TARGETARCH_ARM_SUPPORTS_SRAMV1
  // Format 1 nicht unterstützt
  pRamAdr := 0$^XRamCell;
#endif

END_FUNCTION // Add_sRam_I
#else
FUNCTION AWL Add_sRam_I
VAR_INPUT
	CRC32		: UDINT;
END_VAR
VAR_OUTPUT
	pRamAdr		: ^XramCell;
END_VAR
VAR
   RamStart     : ^XramHdr;
END_VAR
		l.d			pRamAdr,0
 		L.EDI 		_S_RAM_Hptr
 		L.EDI		(EDI+MRAM_DESCR.DataStart)
		S.EDI		RamStart

		// Die folgende Schleife geht die Verkettung der XRAM-Blöcke durch
		// bis das Ende erreicht ist. Am Ende zeigt EBX auf

SearchLoop
		L.EDX     	(EDI+XRAMHDR.udEntries)

		// Abbruch, wenn ein XRAM-Block weniger als 500 XRAM-Zellen enthält
		CMP.EDX		X_RAM_CELLS
		JNE			TheEnd

		// Abbruch, wenn kein Zeiger auf einen weiteren XRAM-Block existiert
		CMP.D		(EDI + XRAMHDR.aData[0] + SIZEOF(XRamCell)*X_RAM_CELLS + XRamCell.udCRC32),1954
		JNE			TheEnd

		// offset zum nächsten block
   		L.EDI		(EDI + XRAMHDR.aData[0] + SIZEOF(XRamCell)*X_RAM_CELLS + XRamCell.udData)
   		ADD.EDI 	RamStart
   		JMP			SearchLoop

TheEnd
		IMUL.EBX	EDX, SIZEOF(XRamCell)
   		ADD.EBX		XRAMHDR.aData[0]

// There is Place in our list, Write It

		CMP.EBX		XRAMHDR.aData[X_RAM_CELLS]
		JNE			MakeNewEntry

// Neuen Block anlegen  und eintragen

		L.EAX		EDI				// pointer auf letzte zelle
		ADD.EAX		EBX

		PUSH		EAX				// place for result
		PUSH		EAX				// Parameter
		CALL		IniNewRamBlock
		POP			EAX				// Parameter
		POP			EAX				// Result

		O.EAX		EAX
		JNZ			GotMemory
		//////////////////////////
		// out of memory !!!    //
		//////////////////////////
		S.EAX		pRamAdr
		L.D			LDR_outOfSramMem, 1     // im Flag merken, dass keine Sram-Speicher mehr vorhanden ist
		JMP			Add_sRam_I_END

GotMemory
		PUSHAD
		CALL		GET_USED_S_RAM	// Memory updaten
		POPAD

		L.EDI		RamStart
		ADD.EDI		EAX

		L.EAX		CRC32
		L.EBX		XRAMHDR.aData[0]

//------------------------------------------------------
// Block belegen und auf ungültig setzen
//------------------------------------------------------

MakeNewEntry

		S.EAX		(EDI+EBX+XRamCell.udCRC32)
		L.D			(EDI+EBX+XRamCell.udData),0
		S.EAX		(EDI+EBX+XRamCell.udChk)

		L.D			(EDI+EBX+XRamCell.udType),16#00000000  // Type = RAM,Daten nicht gültig

		L.ECX		(EDI+XRAMHDR.udEntries)
		INC			ECX
		S.ECX		(EDI+XRAMHDR.udEntries)
		NOT			ECX
		S.ECX		(EDI+XRAMHDR.udChk)

		// --- Pointer auf Zelle Mitgeben ---

		L.EAX		EDI
		ADD.EAX		EBX
		S.EAX		pRamAdr

Add_sRam_I_END

END_FUNCTION // Add_sRam_I
#endif

//---------------------------------------------
// im neuen ram die verbindung zum s-ram suchen
//---------------------------------------------
// Wird von allen S-Ram klassen verwendet um das objekt mit den
// Daten zu verbinden

// auch mit Erweiterung wissen wir ob es ein RAMex ist anhand der Kennung oder nicht

#ifdef _LSL_TARGETARCH_ARM
FUNCTION Find_sRam_I
VAR_INPUT
#pragma warning(disable:73)
	_S_RAM_Hptr0: ^MRAM_DESCR;
	CRC32		: UDINT;
#pragma warning(default:73)
END_VAR
VAR_OUTPUT
	pRamAdr		: ^XramCell;
END_VAR
#ifdef _LSL_TARGETARCH_ARM_SUPPORTS_SRAMV1
VAR
   RamStart     : ^XramHdr;

   FirstChain   :^XramCell;  // pointer to first chain
   LastFoundNr	:UDINT;

   DirNr		:UDINT;
   DirIndex		:UDINT;

   NewFoundNr	:UDINT;

   pXramHdr     : ^XRAMHDR;
   pXramCell	  :^XramCell;
   nRest        : DINT;
   nLoops       : DINT;
END_VAR

  pRamAdr := 0$^XramCell;
  RamStart := _S_RAM_Hptr0^.DataStart;

//-- Ptr to Cell 500 of first block, where we store the element nr auf the previous RAM object
  FirstChain := #RamStart^.aData[X_RAM_CELLS];

// convert Nr into list + index
  LastFoundNr := FirstChain^.udType AND 16#Fffff;

// spezial situation if the first Objekt and List ist empty
  IF (LastFoundNr = 0) & (RamStart^.udEntries = 0) THEN
    RETURN;
  END_IF;

// Select startingPoint by getting the right list + Index
  DirNr := LastFoundNr / X_RAM_CELLS;
  DirIndex := LastFoundNr MOD X_RAM_CELLS;

//-- Liste suchen (über verkettung)--
  pXramHdr := RamStart;
  WHILE DirNr > 0 DO
    pXramHdr := RamStart + pXramHdr^.aData[X_RAM_CELLS].udData; // offset zum nächsten block
    DirNr -= 1;
  END_WHILE;
// -- index suchen  -
  pXramCell := #pXramHdr^.aData[DirIndex];

  nRest := pXramHdr^.udEntries$DINT - DirIndex$DINT;
  IF nRest < 0 THEN
    // wenn bei der Subtraktion eine neg.Zahl rauskommt, dann stimmen die Daten im Sram nicht
    RETURN;
  END_IF;

  NewFoundNr := LastFoundNr;
  IF LastFoundNr = 0 THEN
    // nr 0 suchen wir von vorne
    nLoops := 1;
  ELSE
    // zuerst von LastFoundNr bis ende, dann von vorne suchen
    nLoops := 2;
  END_IF;

  WHILE nLoops > 0 DO
    WHILE nRest > 0 DO

      WHILE nRest > 0 DO
        NewFoundNr += 1;
        pXramCell += SIZEOF(XRamCell);
        nRest -= 1;
        IF CRC32 = pXramCell^.udCRC32 THEN
          // gefunden
          FirstChain^.udType := RamValid OR NewFoundNr; // memorize where we are now to make search faster
          pRamAdr := pXramCell;
          RETURN;
        END_IF;
      END_WHILE;

      // See if there is another list
      IF pXramCell^.udCRC32 = 1954 THEN
        pXramHdr := RamStart + pXramHdr^.aData[X_RAM_CELLS].udData; // offset zum nächsten block
        nRest := pXramHdr^.udEntries$DINT;
      END_IF;

    END_WHILE;

    // Zweiter Schleifendurchlauf von vorne
    pXramHdr := RamStart;
    pXramCell := #pXramHdr^.aData[0];
    nLoops -= 1;

  END_WHILE;
#else // _LSL_TARGETARCH_ARM_SUPPORTS_SRAMV1
  pRamAdr := 0$^XramCell;
#endif

END_FUNCTION // Find_sRam_I
#else
FUNCTION AWL Find_sRam_I
VAR_INPUT
	_S_RAM_Hptr0: ^MRAM_DESCR;
	CRC32		: UDINT;
END_VAR
VAR_OUTPUT
	pRamAdr		: ^XramCell;
END_VAR
VAR
   RamStart     : ^XramHdr;

   FirstChain   :^XramCell;  // pointer to first chain
   LastFoundNr	:UDINT;

   DirNr		:UDINT;
   Dirindex		:UDINT;

   LastListAdr	:^XramHdr;  // Memory for end of list
   LastEleOffs	:^XramCell;
   NewFoundNr	:UDINT;

END_VAR
		l.d			pRamAdr,0
   		L.EDI 		_S_RAM_Hptr0
		L.EAX		(EDI+MRAM_DESCR.DataValid)

   		L.EDI		(EDI+MRAM_DESCR.DataStart)
		S.EDI		RamStart

//-- Ptr to Cell 500 of first block, where we store the element nr auf the previous RAM object

		L.EBX		EDI
		ADD.EBX		XRAMHDR.aData[X_RAM_CELLS]
		S.EBX		FirstChain

// convert Nr into list + index

		L.EAX		(EBX+xRamCell.udType)
		A.EAX		16#Fffff
		S.EAX		LastFoundNr

// spezial situation if the first Objekt and List ist empty

		JNZ			ItIsNotTheFirst
		CMP.D		(EDI+XRAMHDR.udEntries),0
		Jne			ItIsNotTheFirst
		JMP			Find_sRam_I_END

// Select startingPoint by getting the right list + Index

ItIsNotTheFirst

		CLR			EDX
		L.ECX		X_RAM_CELLS
		DIV			ECX
		S.EAX		DirNr
		S.EDX		DirIndex

//-- Liste suchen (über verkettung)--

		O.EAX		EAX
		JZ			Go1
SFLP
   		L.EDI		(EDI+XRAMHDR.aData[X_RAM_CELLS].udData) 	  // offset zum nächsten block
   		ADD.EDI 	RamStart
		DEC			EAX
		JNZ			SFLP

// -- index suchen (ist rest der division) -

Go1		IMUL.EBX	EDX,SIZEOF(XRamCell)
   		ADD.EBX		XRAMHDR.aData[0]

//-------------------------------
// -- Von Jetzt bis ende suchen--
//-------------------------------

//  EDX = INDEX In LISTE

		L.ECX		(EDI+XRAMHDR.udEntries)//EDI:blockPtr
		SUB.ECX		EDX//EDX:DirIndex
    JC      ItsNotInTheList // wenn bei der Subtraktion eine neg.Zahl rauskommt, dann stimmen die Daten im Sram nicht
   		L.EAX		CRC32

		L.EDX        LastFoundNr
		O.EDX		EDX						// nr 0 suchen wir von vorne
		JZ			SearchToEndLoop

		INC			EDX						// NewFoundNr ab dann immer den nächsten
		ADD.EBX  	SIZEOF(XRamCell)
		LOOP	 	SearchToEndLoop			//--> Suchen, ECX:rest.Anz.Entries im Block

		JMP			SearchToEnd_X

SearchToEndLoop

		CMP.EAX		(EDI+EBX+XRamCell.udCRC32)
		JE			RamFound
		INC			EDX						// NewFoundNr
		ADD.EBX  	SIZEOF(XRamCell)
		LOOP	 	SearchToEndLoop			//--> Suchen
SearchToEnd_X
		CMP.EBX		XRAMHDR.aData[X_RAM_CELLS]
		JNE			NoMatchAtEnd

// See if there is another list

   		CMP.D		(EDI+EBX+XRamCell.udCRC32),1954
		JNE			NoMatchAtEnd

   		L.EDI		(EDI+EBX+XRamCell.udData) 	  // offset zum nächsten block
   		ADD.EDI 	RamStart
		L.ECX		(EDI+XRAMHDR.udEntries)
  		L.EBX		XRAMHDR.aData[0]
   		JMP			SearchToEndLoop

// We are at the end and found no entry

NoMatchAtEnd

   		S.EDI		LastListAdr	 // Memory for end of list
   		S.EBX		LastEleOffs
		S.EDX		NewFoundNr

//----------------------------
// now we search from beginning
//-----------------------------

		CLR			EDX   // 		 	NewFoundNr
		L.EDI		RamStart

		L.ECX		(EDI+XRAMHDR.udEntries)
   		L.EBX		XRAMHDR.aData[0]

SearchFromBegLoop

  		CMP.EAX		(EDI+EBX+XRamCell.udCRC32)
   		Je			RamFound

		INC			EDX
		ADD.EBX  	SIZEOF(XRamCell)
		LOOP	 	SearchFromBegLoop		//--> Suchen

		CMP.EBX		XRAMHDR.aData[X_RAM_CELLS]
		JNE			ItsNotInTheList

// See if there is another list

   		CMP.D		(EDI+EBX+XRamCell.udCRC32),1954
		JNE			ItsNotInTheList

   		L.EDI		(EDI+EBX+XRamCell.udData) 	  // offset zum nächsten block
   		ADD.EDI 	RamStart
		L.ECX		(EDI+XRAMHDR.udEntries)
   		L.EBX		XRAMHDR.aData[0]

   		JMP			SearchFromBegLoop

//---------------------------------------------------
// Now we definately know that this is an new element
//---------------------------------------------------

ItsNotInTheList
		JMP			Find_sRam_I_END

// --- Gefunden, Pointer auf Zelle Mitgeben ---

RamFound

// memorize where we are now to make search faster

		L.EAX		FirstChain
		O.EDX		RamValid
		S.EDX		(EAX+xRamCell.udType)

   		L.EAX		EDI
		ADD.EAX		EBX
   		S.EAX		pRamAdr
